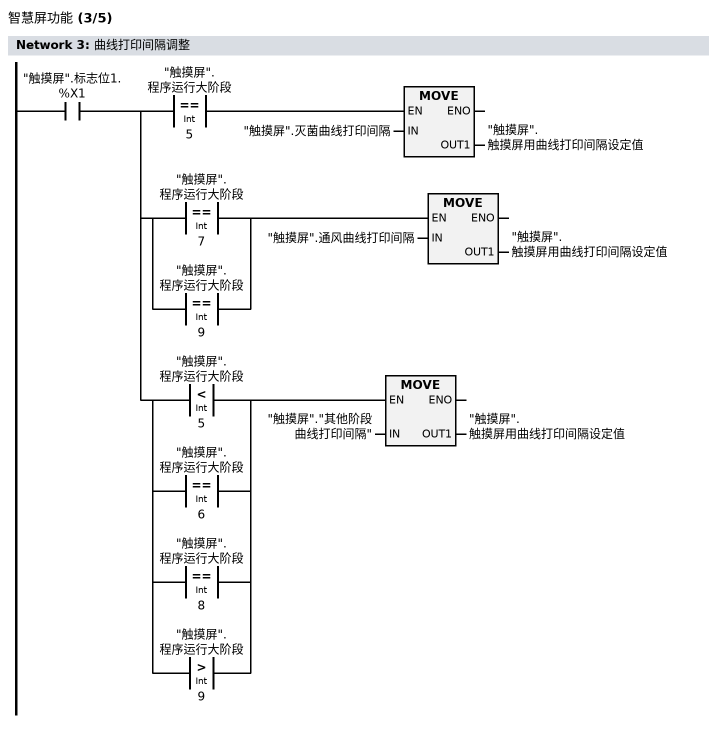
   RUNG wire#powerrail
      Contact( "触摸屏".标志位1.%X1 )
      wire#w1
      { S7_Templates := "SrcType := Int" } EQ_Contact(in1 := "触摸屏".程序运行大阶段, in2 := 5)
      Move(in := "触摸屏".灭菌曲线打印间隔, out1 => "触摸屏".触摸屏用曲线打印间隔设定值)
   END_RUNG
   RUNG wire#w1
      { S7_Templates := "SrcType := Int" } EQ_Contact(in1 := "触摸屏".程序运行大阶段, in2 := 7)
      wire#w2
      Move(in := "触摸屏".通风曲线打印间隔, out1 => "触摸屏".触摸屏用曲线打印间隔设定值)
   END_RUNG
   RUNG wire#w1
      { S7_Templates := "SrcType := Int" } EQ_Contact(in1 := "触摸屏".程序运行大阶段, in2 := 9)
   END_RUNG wire#w2
   RUNG wire#w1
      { S7_Templates := "SrcType := Int" } LT_Contact(in1 := "触摸屏".程序运行大阶段, in2 := 5)
      wire#w3
      Move(in := "触摸屏"."其他阶段 曲线打印间隔", out1 => "触摸屏".触摸屏用曲线打印间隔设定值)
   END_RUNG
   RUNG wire#w1
      { S7_Templates := "SrcType := Int" } EQ_Contact(in1 := "触摸屏".程序运行大阶段, in2 := 6)
   END_RUNG wire#w3
   RUNG wire#w1
      { S7_Templates := "SrcType := Int" } EQ_Contact(in1 := "触摸屏".程序运行大阶段, in2 := 8)
   END_RUNG wire#w3
   RUNG wire#w1
      { S7_Templates := "SrcType := Int" } GT_Contact(in1 := "触摸屏".程序运行大阶段, in2 := 9)
   END_RUNG wire#w3
   // the same network as SCL:
   IF "触摸屏".标志位1.%X1 AND ("触摸屏".程序运行大阶段 = 5) THEN "触摸屏".触摸屏用曲线打印间隔设定值 := "触摸屏".灭菌曲线打印间隔; END_IF;
   IF "触摸屏".标志位1.%X1 AND (("触摸屏".程序运行大阶段 = 7) OR ("触摸屏".程序运行大阶段 = 9)) THEN
       "触摸屏".触摸屏用曲线打印间隔设定值 := "触摸屏".通风曲线打印间隔;
   END_IF;
   IF "触摸屏".标志位1.%X1 AND (("触摸屏".程序运行大阶段 < 5) OR ("触摸屏".程序运行大阶段 = 6) OR ("触摸屏".程序运行大阶段 = 8) OR ("触摸屏".程序运行大阶段 > 9)) THEN
       "触摸屏".触摸屏用曲线打印间隔设定值 := "触摸屏"."其他阶段 曲线打印间隔";
   END_IF;
END_REGION

REGION Network 4: 报表打印控制 报表间隔控制，printflag， "DB48.DBD684", 用于控制报表打印
   // 曲线间隔：灭菌20秒，通风60秒，其他10秒
   // 报表间隔：1：预处理  10分钟
   // 2：保压   10分钟
   // 3：加湿    10分钟
   // 4：加药    10分钟
   // 5：灭菌    20分钟
   // 6：脉动    10分钟
   // 7：通风   60分钟
   // 8：紧急脉动 10分钟
   // 9：紧急通风  30分钟
   // 10：结束
   // 
   // 智慧屏曲线打印会打印：大阶段 小阶段  printflag+定时存储的数据，定时存储需要再global全局设置
   //             报表打印会打印：大阶段 小阶段  printflag
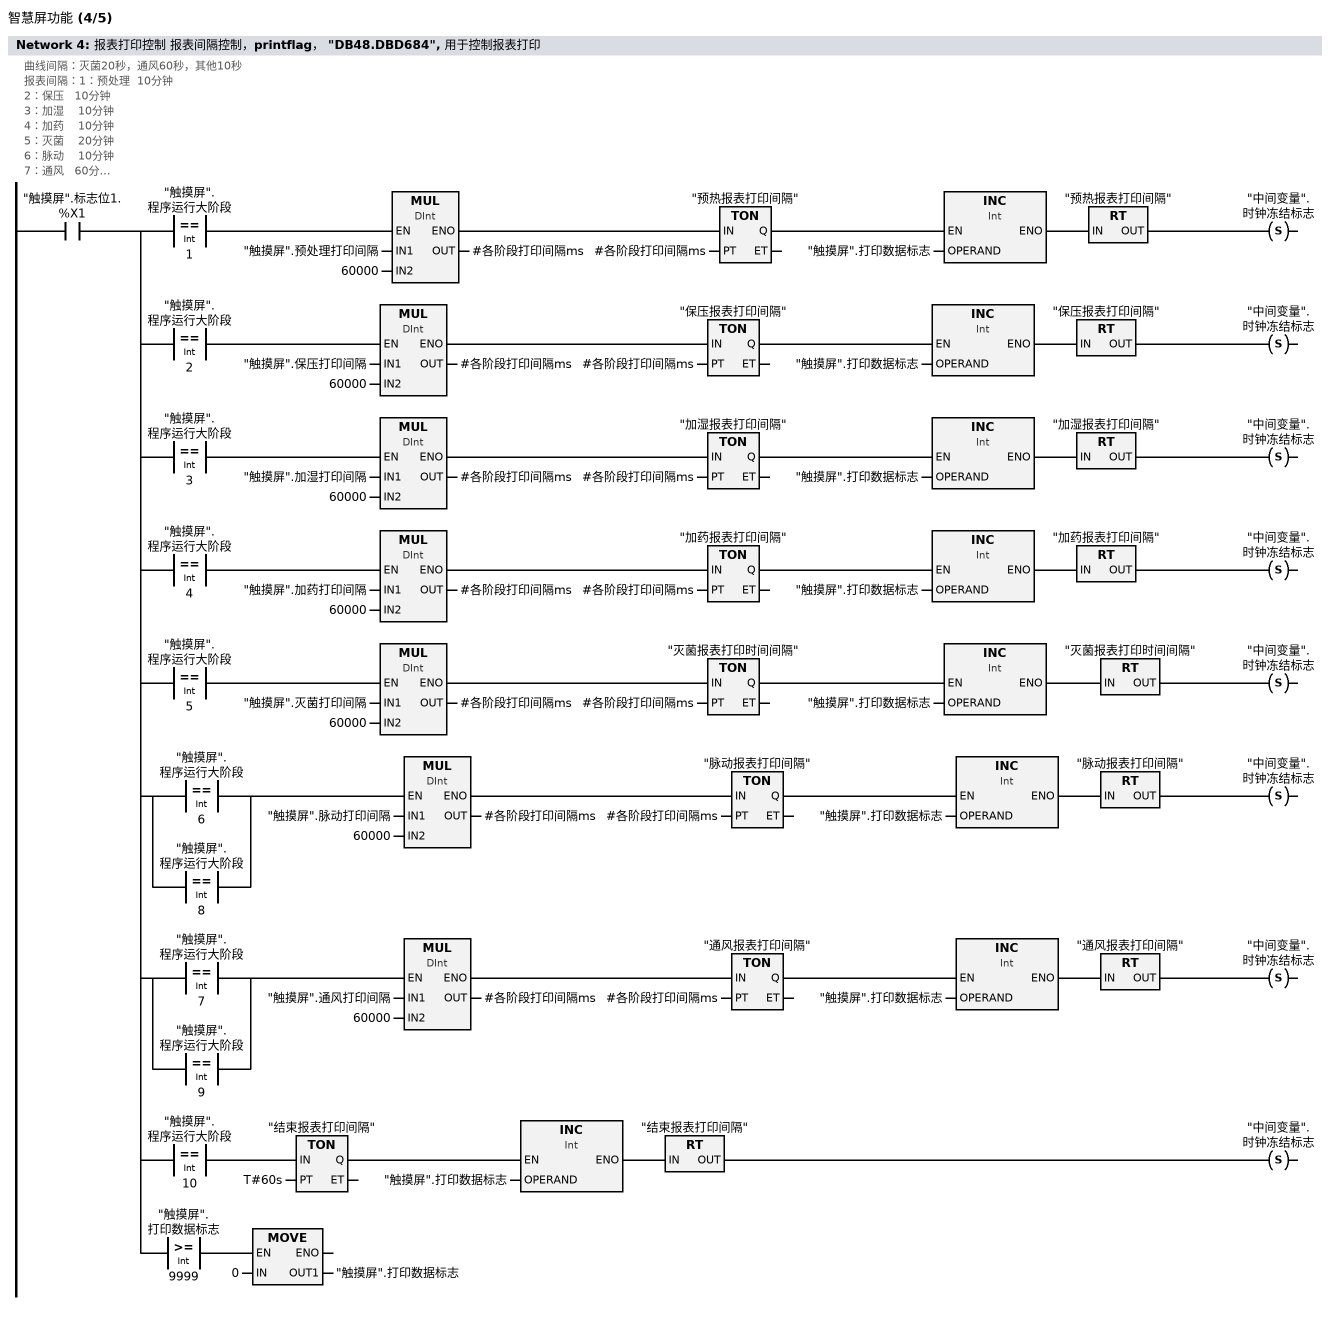
   #_w1 := "触摸屏".标志位1.%X1 AND ("触摸屏".程序运行大阶段 = 1);
   IF #_w1 THEN #各阶段打印间隔ms := "触摸屏".预处理打印间隔 * 60000; END_IF;
   "预热报表打印间隔".TON(IN := #_w1, PT := #各阶段打印间隔ms);
   IF "预热报表打印间隔".Q THEN "触摸屏".打印数据标志 := "触摸屏".打印数据标志 + 1; END_IF;
   #_w2 := "预热报表打印间隔".Q;
   IF #_w2 THEN
       RESET_TIMER("预热报表打印间隔");
       "中间变量".时钟冻结标志 := TRUE;
   END_IF;
   #_w3 := "触摸屏".标志位1.%X1 AND ("触摸屏".程序运行大阶段 = 2);
   IF #_w3 THEN #各阶段打印间隔ms := "触摸屏".保压打印间隔 * 60000; END_IF;
   "保压报表打印间隔".TON(IN := #_w3, PT := #各阶段打印间隔ms);
   IF "保压报表打印间隔".Q THEN "触摸屏".打印数据标志 := "触摸屏".打印数据标志 + 1; END_IF;
   #_w4 := "保压报表打印间隔".Q;
   IF #_w4 THEN
       RESET_TIMER("保压报表打印间隔");
       "中间变量".时钟冻结标志 := TRUE;
   END_IF;
   #_w5 := "触摸屏".标志位1.%X1 AND ("触摸屏".程序运行大阶段 = 3);
   IF #_w5 THEN #各阶段打印间隔ms := "触摸屏".加湿打印间隔 * 60000; END_IF;
   "加湿报表打印间隔".TON(IN := #_w5, PT := #各阶段打印间隔ms);
   IF "加湿报表打印间隔".Q THEN "触摸屏".打印数据标志 := "触摸屏".打印数据标志 + 1; END_IF;
   #_w6 := "加湿报表打印间隔".Q;
   IF #_w6 THEN
       RESET_TIMER("加湿报表打印间隔");
       "中间变量".时钟冻结标志 := TRUE;
   END_IF;
   #_w7 := "触摸屏".标志位1.%X1 AND ("触摸屏".程序运行大阶段 = 4);
   IF #_w7 THEN #各阶段打印间隔ms := "触摸屏".加药打印间隔 * 60000; END_IF;
   "加药报表打印间隔".TON(IN := #_w7, PT := #各阶段打印间隔ms);
   IF "加药报表打印间隔".Q THEN "触摸屏".打印数据标志 := "触摸屏".打印数据标志 + 1; END_IF;
   #_w8 := "加药报表打印间隔".Q;
   IF #_w8 THEN
       RESET_TIMER("加药报表打印间隔");
       "中间变量".时钟冻结标志 := TRUE;
   END_IF;
   #_w9 := "触摸屏".标志位1.%X1 AND ("触摸屏".程序运行大阶段 = 5);
   IF #_w9 THEN #各阶段打印间隔ms := "触摸屏".灭菌打印间隔 * 60000; END_IF;
   "灭菌报表打印时间间隔".TON(IN := #_w9, PT := #各阶段打印间隔ms);
   IF "灭菌报表打印时间间隔".Q THEN "触摸屏".打印数据标志 := "触摸屏".打印数据标志 + 1; END_IF;
   #_w10 := "灭菌报表打印时间间隔".Q;
   IF #_w10 THEN
       RESET_TIMER("灭菌报表打印时间间隔");
       "中间变量".时钟冻结标志 := TRUE;
   END_IF;
   #_w11 := "触摸屏".标志位1.%X1 AND (("触摸屏".程序运行大阶段 = 6) OR ("触摸屏".程序运行大阶段 = 8));
   IF #_w11 THEN #各阶段打印间隔ms := "触摸屏".脉动打印间隔 * 60000; END_IF;
   "脉动报表打印间隔".TON(IN := #_w11, PT := #各阶段打印间隔ms);
   IF "脉动报表打印间隔".Q THEN "触摸屏".打印数据标志 := "触摸屏".打印数据标志 + 1; END_IF;
   #_w12 := "脉动报表打印间隔".Q;
   IF #_w12 THEN
       RESET_TIMER("脉动报表打印间隔");
       "中间变量".时钟冻结标志 := TRUE;
   END_IF;
   #_w13 := "触摸屏".标志位1.%X1 AND (("触摸屏".程序运行大阶段 = 7) OR ("触摸屏".程序运行大阶段 = 9));
   IF #_w13 THEN #各阶段打印间隔ms := "触摸屏".通风打印间隔 * 60000; END_IF;
   "通风报表打印间隔".TON(IN := #_w13, PT := #各阶段打印间隔ms);
   IF "通风报表打印间隔".Q THEN "触摸屏".打印数据标志 := "触摸屏".打印数据标志 + 1; END_IF;
   #_w14 := "通风报表打印间隔".Q;
   IF #_w14 THEN
       RESET_TIMER("通风报表打印间隔");
       "中间变量".时钟冻结标志 := TRUE;
   END_IF;
   "结束报表打印间隔".TON(IN := "触摸屏".标志位1.%X1 AND ("触摸屏".程序运行大阶段 = 10), PT := T#60s);
   IF "结束报表打印间隔".Q THEN "触摸屏".打印数据标志 := "触摸屏".打印数据标志 + 1; END_IF;
   #_w15 := "结束报表打印间隔".Q;
   IF #_w15 THEN
       RESET_TIMER("结束报表打印间隔");
       "中间变量".时钟冻结标志 := TRUE;
   END_IF;
   IF "触摸屏".标志位1.%X1 AND ("触摸屏".打印数据标志 >= 9999) THEN "触摸屏".打印数据标志 := 0; END_IF;
END_REGION

REGION Network 5: 冻结PLC时钟标志，为了智慧屏能获取 阶段变化的真实时间，阶段变化后需要冻结PLC时间2秒钟
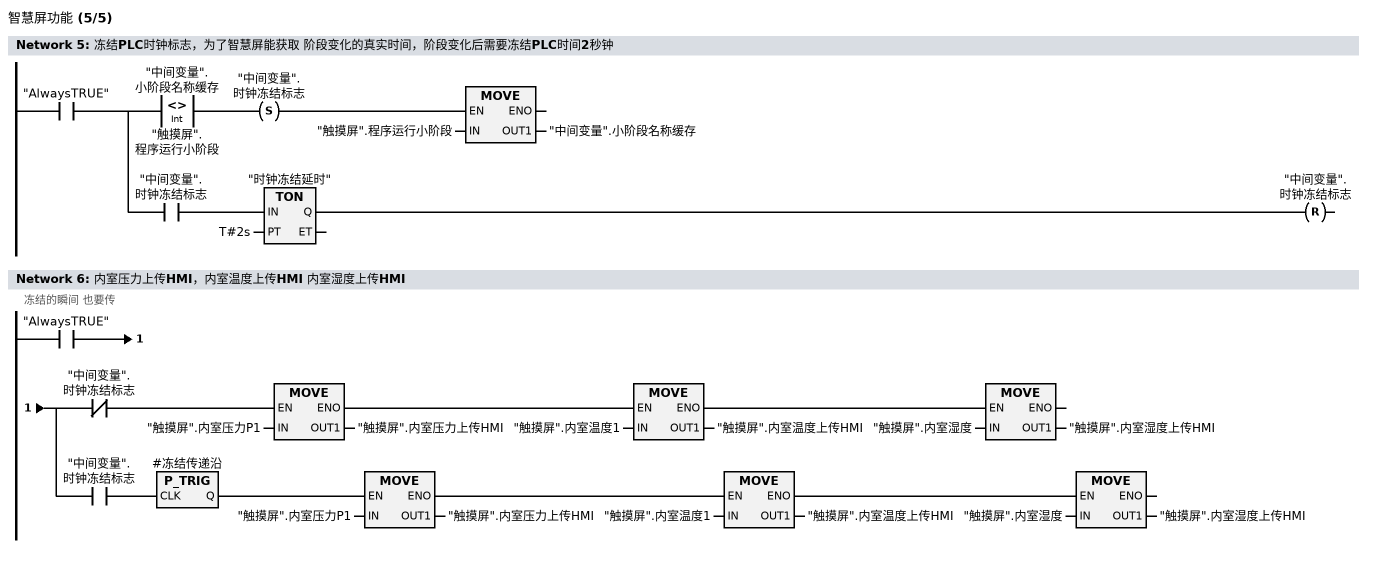
   IF "AlwaysTRUE" AND ("中间变量".小阶段名称缓存 <> "触摸屏".程序运行小阶段) THEN
       "中间变量".时钟冻结标志 := TRUE;
       "中间变量".小阶段名称缓存 := "触摸屏".程序运行小阶段;
   END_IF;
   "时钟冻结延时".TON(IN := "AlwaysTRUE" AND "中间变量".时钟冻结标志, PT := T#2s);
   IF "时钟冻结延时".Q THEN "中间变量".时钟冻结标志 := FALSE; END_IF;
END_REGION

REGION Network 6: 内室压力上传HMI，内室温度上传HMI 内室湿度上传HMI
   // 冻结的瞬间 也要传
   RUNG wire#powerrail
      Contact( "AlwaysTRUE" )
      wire#w1
      I_Contact( "中间变量".时钟冻结标志 )
      Move(in := "触摸屏".内室压力P1, out1 => "触摸屏".内室压力上传HMI)
      Move(in := "触摸屏".内室温度1, out1 => "触摸屏".内室温度上传HMI)
      Move(in := "触摸屏".内室湿度, out1 => "触摸屏".内室湿度上传HMI)
   END_RUNG
   RUNG wire#w1
      Contact( "中间变量".时钟冻结标志 )
      P_Trig( #冻结传递沿 )
      Move(in := "触摸屏".内室压力P1, out1 => "触摸屏".内室压力上传HMI)
      Move(in := "触摸屏".内室温度1, out1 => "触摸屏".内室温度上传HMI)
      Move(in := "触摸屏".内室湿度, out1 => "触摸屏".内室湿度上传HMI)
   END_RUNG
   // the same network as SCL:
   IF "AlwaysTRUE" AND NOT "中间变量".时钟冻结标志 THEN
       "触摸屏".内室压力上传HMI := "触摸屏".内室压力P1;
       "触摸屏".内室温度上传HMI := "触摸屏".内室温度1;
       "触摸屏".内室湿度上传HMI := "触摸屏".内室湿度;
   END_IF;
   #_w1 := "AlwaysTRUE" AND "中间变量".时钟冻结标志;
   #_w2 := #_w1 AND NOT #冻结传递沿;   // rising edge
   #冻结传递沿 := #_w1;
   IF #_w2 THEN
       "触摸屏".内室压力上传HMI := "触摸屏".内室压力P1;
       "触摸屏".内室温度上传HMI := "触摸屏".内室温度1;
       "触摸屏".内室湿度上传HMI := "触摸屏".内室湿度;
   END_IF;
END_REGION
END_FUNCTION_BLOCK

// folder: 6系统设置

FUNCTION_BLOCK "系统参数设置"   // FB21, LAD
{ S7_Optimized_Access := 'TRUE' }
VERSION : 0.1
   VAR
      催化剂使用时间秒 : Int;
      催化剂使用时间分 : Int;
      催化剂使用时间时 : Int;
      催化剂使用统计沿 : Bool;
   END_VAR
   VAR RETAIN
      催化剂使用统计秒 : Int;
   END_VAR
   VAR_TEMP
      中间变量 : Int;
   END_VAR
   VAR_TEMP   // added for the SCL form of the ladder/FBD networks
      _w1 : Bool;
      _w2 : Bool;
   END_VAR
BEGIN

REGION Network 1: 解毒阀开启时间统计，即催化剂使用时间统计
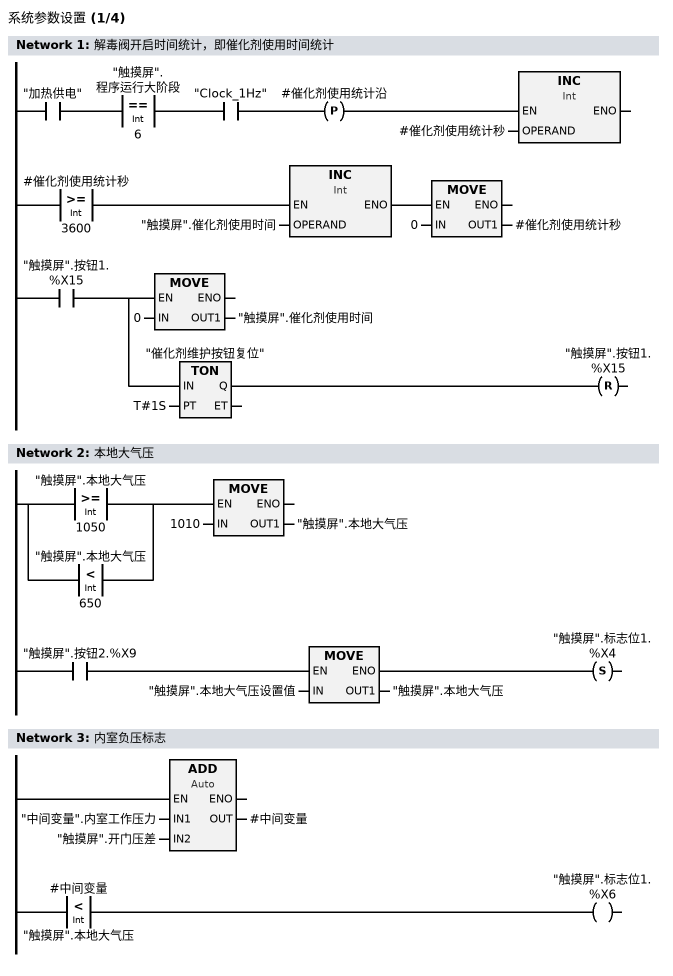
   #_w1 := "加热供电" AND ("触摸屏".程序运行大阶段 = 6) AND "Clock_1Hz";
   #_w2 := #_w1 AND NOT #催化剂使用统计沿;   // rising edge
   #催化剂使用统计沿 := #_w1;
   IF #_w2 THEN #催化剂使用统计秒 := #催化剂使用统计秒 + 1; END_IF;
   IF #催化剂使用统计秒 >= 3600 THEN
       "触摸屏".催化剂使用时间 := "触摸屏".催化剂使用时间 + 1;
       #催化剂使用统计秒 := 0;
   END_IF;
   IF "触摸屏".按钮1.%X15 THEN "触摸屏".催化剂使用时间 := 0; END_IF;
   "催化剂维护按钮复位".TON(IN := "触摸屏".按钮1.%X15, PT := T#1S);
   IF "催化剂维护按钮复位".Q THEN "触摸屏".按钮1.%X15 := FALSE; END_IF;
END_REGION

REGION Network 2: 本地大气压
   RUNG wire#powerrail
      { S7_Templates := "SrcType := Int" } GE_Contact(in1 := "触摸屏".本地大气压, in2 := 1050)
      wire#w1
      Move(in := 1010, out1 => "触摸屏".本地大气压)
   END_RUNG
   RUNG wire#powerrail
      { S7_Templates := "SrcType := Int" } LT_Contact(in1 := "触摸屏".本地大气压, in2 := 650)
   END_RUNG wire#w1
   RUNG wire#powerrail
      Contact( "触摸屏".按钮2.%X9 )
      Move(in := "触摸屏".本地大气压设置值, out1 => "触摸屏".本地大气压)
      S_Coil( "触摸屏".标志位1.%X4 )
   END_RUNG
   // the same network as SCL:
   IF ("触摸屏".本地大气压 >= 1050) OR ("触摸屏".本地大气压 < 650) THEN "触摸屏".本地大气压 := 1010; END_IF;
   IF "触摸屏".按钮2.%X9 THEN
       "触摸屏".本地大气压 := "触摸屏".本地大气压设置值;
       "触摸屏".标志位1.%X4 := TRUE;
   END_IF;
END_REGION

REGION Network 3: 内室负压标志
   RUNG wire#powerrail
      Add(in1 := "中间变量".内室工作压力, in2 := "触摸屏".开门压差, out => #中间变量)
   END_RUNG
   RUNG wire#powerrail
      { S7_Templates := "SrcType := Int" } LT_Contact(in1 := #中间变量, in2 := "触摸屏".本地大气压)
      Coil( "触摸屏".标志位1.%X6 )
   END_RUNG
   // the same network as SCL:
   #中间变量 := "中间变量".内室工作压力 + "触摸屏".开门压差;
   "触摸屏".标志位1.%X6 := #中间变量 < "触摸屏".本地大气压;
END_REGION

REGION Network 4: 蜂鸣器参数
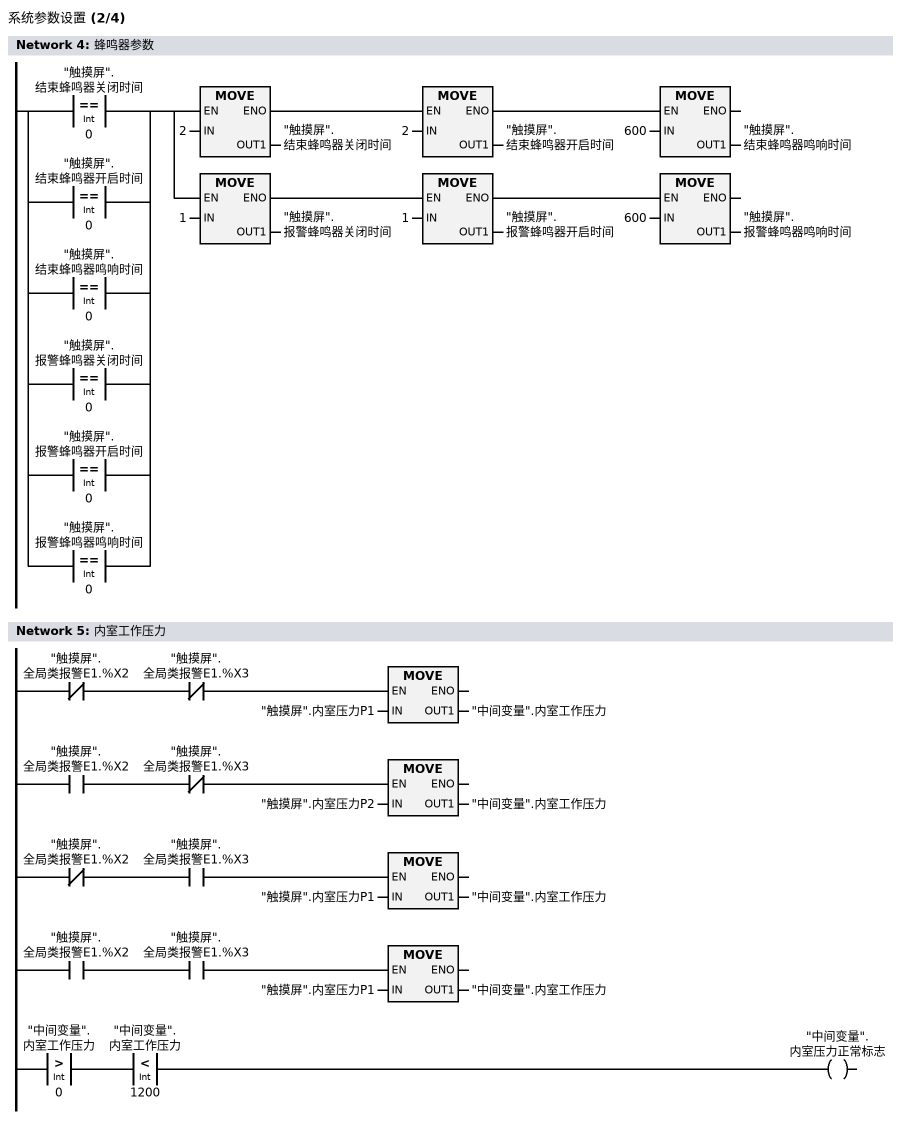
   RUNG wire#powerrail
      { S7_Templates := "SrcType := Int" } EQ_Contact(in1 := "触摸屏".结束蜂鸣器关闭时间, in2 := 0)
      wire#w1
      Move(in := 2, out1 => "触摸屏".结束蜂鸣器关闭时间)
      Move(in := 2, out1 => "触摸屏".结束蜂鸣器开启时间)
      Move(in := 600, out1 => "触摸屏".结束蜂鸣器鸣响时间)
   END_RUNG
   RUNG wire#powerrail
      { S7_Templates := "SrcType := Int" } EQ_Contact(in1 := "触摸屏".结束蜂鸣器开启时间, in2 := 0)
   END_RUNG wire#w1
   RUNG wire#powerrail
      { S7_Templates := "SrcType := Int" } EQ_Contact(in1 := "触摸屏".结束蜂鸣器鸣响时间, in2 := 0)
   END_RUNG wire#w1
   RUNG wire#powerrail
      { S7_Templates := "SrcType := Int" } EQ_Contact(in1 := "触摸屏".报警蜂鸣器关闭时间, in2 := 0)
   END_RUNG wire#w1
   RUNG wire#powerrail
      { S7_Templates := "SrcType := Int" } EQ_Contact(in1 := "触摸屏".报警蜂鸣器开启时间, in2 := 0)
   END_RUNG wire#w1
   RUNG wire#powerrail
      { S7_Templates := "SrcType := Int" } EQ_Contact(in1 := "触摸屏".报警蜂鸣器鸣响时间, in2 := 0)
   END_RUNG wire#w1
   RUNG wire#w1
      Move(in := 1, out1 => "触摸屏".报警蜂鸣器关闭时间)
      Move(in := 1, out1 => "触摸屏".报警蜂鸣器开启时间)
      Move(in := 600, out1 => "触摸屏".报警蜂鸣器鸣响时间)
   END_RUNG
   // the same network as SCL:
   #_w1 := ("触摸屏".结束蜂鸣器关闭时间 = 0) OR ("触摸屏".结束蜂鸣器开启时间 = 0) OR ("触摸屏".结束蜂鸣器鸣响时间 = 0) OR ("触摸屏".报警蜂鸣器关闭时间 = 0) OR ("触摸屏".报警蜂鸣器开启时间 = 0) OR ("触摸屏".报警蜂鸣器鸣响时间 = 0);
   #_w2 := ("触摸屏".结束蜂鸣器关闭时间 = 0) OR ("触摸屏".结束蜂鸣器开启时间 = 0) OR ("触摸屏".结束蜂鸣器鸣响时间 = 0) OR ("触摸屏".报警蜂鸣器关闭时间 = 0) OR ("触摸屏".报警蜂鸣器开启时间 = 0) OR ("触摸屏".报警蜂鸣器鸣响时间 = 0);
   IF #_w2 THEN
       "触摸屏".结束蜂鸣器关闭时间 := 2;
       "触摸屏".结束蜂鸣器开启时间 := 2;
       "触摸屏".结束蜂鸣器鸣响时间 := 600;
   END_IF;
   IF #_w1 THEN
       "触摸屏".报警蜂鸣器关闭时间 := 1;
       "触摸屏".报警蜂鸣器开启时间 := 1;
       "触摸屏".报警蜂鸣器鸣响时间 := 600;
   END_IF;
END_REGION

REGION Network 5: 内室工作压力
   RUNG wire#powerrail
      I_Contact( "触摸屏".全局类报警E1.%X2 )
      I_Contact( "触摸屏".全局类报警E1.%X3 )
      Move(in := "触摸屏".内室压力P1, out1 => "中间变量".内室工作压力)
   END_RUNG
   RUNG wire#powerrail
      Contact( "触摸屏".全局类报警E1.%X2 )
      I_Contact( "触摸屏".全局类报警E1.%X3 )
      Move(in := "触摸屏".内室压力P2, out1 => "中间变量".内室工作压力)
   END_RUNG
   RUNG wire#powerrail
      I_Contact( "触摸屏".全局类报警E1.%X2 )
      Contact( "触摸屏".全局类报警E1.%X3 )
      Move(in := "触摸屏".内室压力P1, out1 => "中间变量".内室工作压力)
   END_RUNG
   RUNG wire#powerrail
      Contact( "触摸屏".全局类报警E1.%X2 )
      Contact( "触摸屏".全局类报警E1.%X3 )
      Move(in := "触摸屏".内室压力P1, out1 => "中间变量".内室工作压力)
   END_RUNG
   RUNG wire#powerrail
      { S7_Templates := "SrcType := Int" } GT_Contact(in1 := "中间变量".内室工作压力, in2 := 0)
      { S7_Templates := "SrcType := Int" } LT_Contact(in1 := "中间变量".内室工作压力, in2 := 1200)
      Coil( "中间变量".内室压力正常标志 )
   END_RUNG
   // the same network as SCL:
   IF NOT "触摸屏".全局类报警E1.%X2 AND NOT "触摸屏".全局类报警E1.%X3 THEN "中间变量".内室工作压力 := "触摸屏".内室压力P1; END_IF;
   IF "触摸屏".全局类报警E1.%X2 AND NOT "触摸屏".全局类报警E1.%X3 THEN "中间变量".内室工作压力 := "触摸屏".内室压力P2; END_IF;
   IF NOT "触摸屏".全局类报警E1.%X2 AND "触摸屏".全局类报警E1.%X3 THEN "中间变量".内室工作压力 := "触摸屏".内室压力P1; END_IF;
   IF "触摸屏".全局类报警E1.%X2 AND "触摸屏".全局类报警E1.%X3 THEN "中间变量".内室工作压力 := "触摸屏".内室压力P1; END_IF;
   "中间变量".内室压力正常标志 := ("中间变量".内室工作压力 > 0) AND ("中间变量".内室工作压力 < 1200);
END_REGION

REGION Network 6: 设备维护
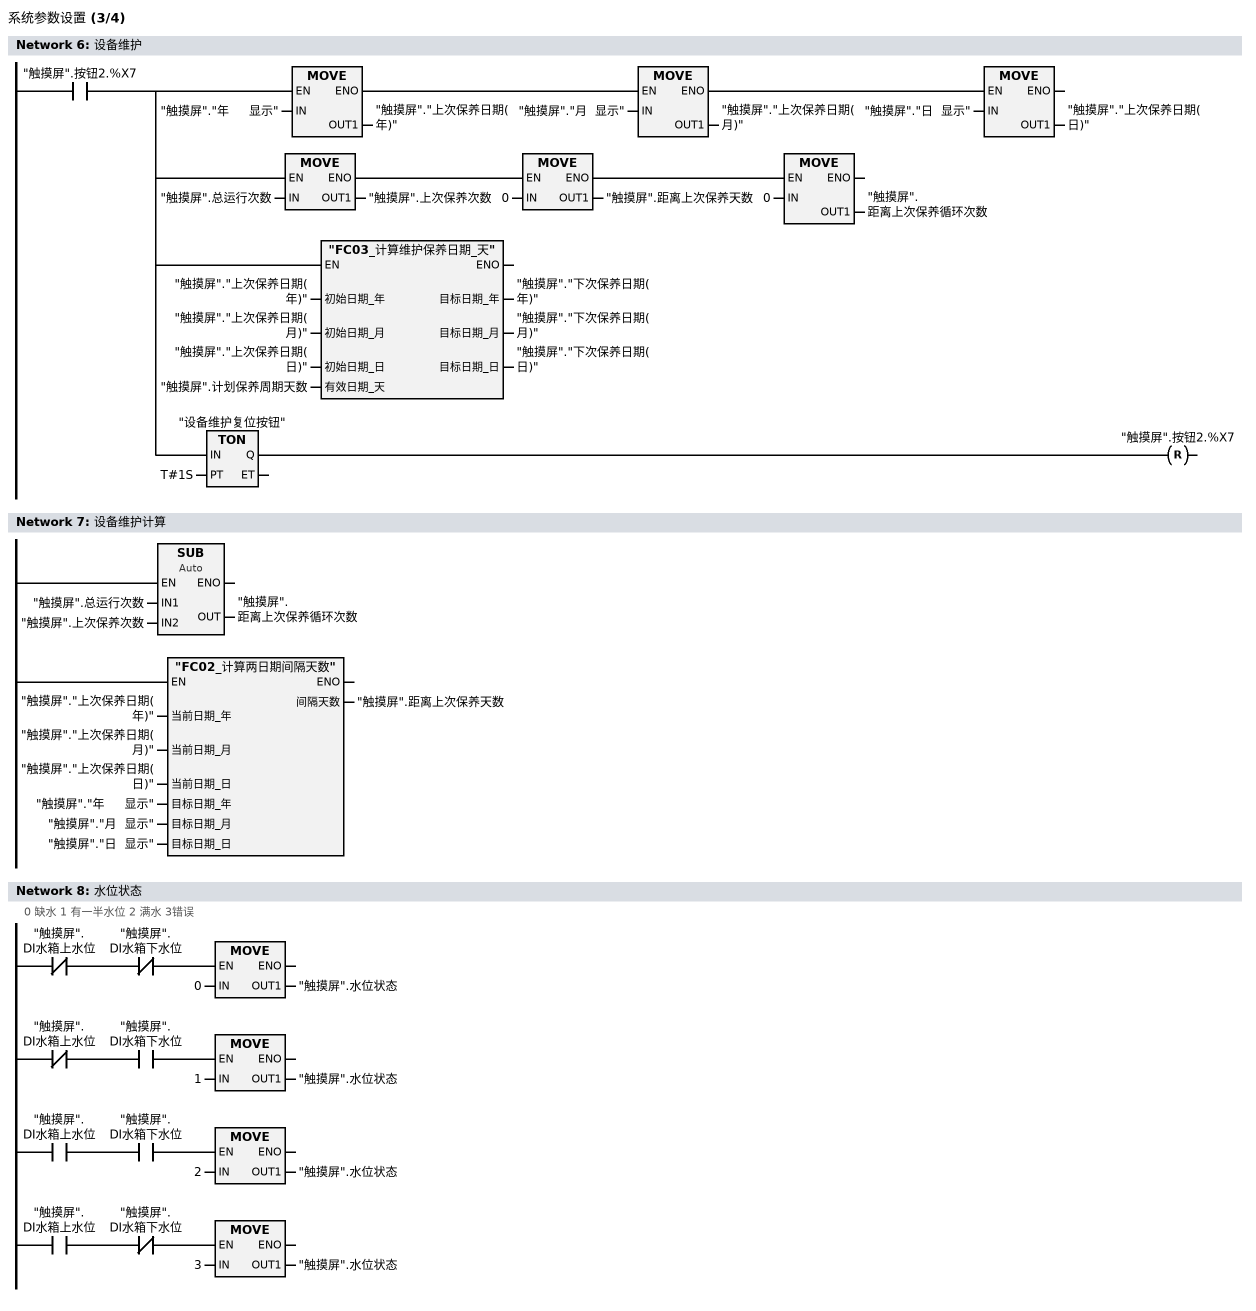
   IF "触摸屏".按钮2.%X7 THEN
       "触摸屏"."上次保养日期(年)" := "触摸屏"."年     显示";
       "触摸屏"."上次保养日期(月)" := "触摸屏"."月  显示";
       "触摸屏"."上次保养日期(日)" := "触摸屏"."日  显示";
       "触摸屏".上次保养次数 := "触摸屏".总运行次数;
       "触摸屏".距离上次保养天数 := 0;
       "触摸屏".距离上次保养循环次数 := 0;
   END_IF;
   #_w1 := "触摸屏".按钮2.%X7;
   IF #_w1 THEN
       "FC03_计算维护保养日期_天"(初始日期_年 := "触摸屏"."上次保养日期(年)",
                         初始日期_月 := "触摸屏"."上次保养日期(月)",
                         初始日期_日 := "触摸屏"."上次保养日期(日)",
                         有效日期_天 := "触摸屏".计划保养周期天数,
                         目标日期_年 => "触摸屏"."下次保养日期(年)",
                         目标日期_月 => "触摸屏"."下次保养日期(月)",
                         目标日期_日 => "触摸屏"."下次保养日期(日)");
   END_IF;
   "设备维护复位按钮".TON(IN := #_w1, PT := T#1S);
   IF "设备维护复位按钮".Q THEN "触摸屏".按钮2.%X7 := FALSE; END_IF;
END_REGION

REGION Network 7: 设备维护计算
   RUNG wire#powerrail
      Sub(in1 := "触摸屏".总运行次数, in2 := "触摸屏".上次保养次数, out => "触摸屏".距离上次保养循环次数)
   END_RUNG
   RUNG wire#powerrail
      "FC02_计算两日期间隔天数"(当前日期_年 := "触摸屏"."上次保养日期(年)", 当前日期_月 := "触摸屏"."上次保养日期(月)", 当前日期_日 := "触摸屏"."上次保养日期(日)", 目标日期_年 := "触摸屏"."年     显示", 目标日期_月 := "触摸屏"."月  显示", 目标日期_日 := "触摸屏"."日  显示", 间隔天数 => "触摸屏".距离上次保养天数)
   END_RUNG
   // the same network as SCL:
   "触摸屏".距离上次保养循环次数 := "触摸屏".总运行次数 - "触摸屏".上次保养次数;
   "FC02_计算两日期间隔天数"(当前日期_年 := "触摸屏"."上次保养日期(年)",
                    当前日期_月 := "触摸屏"."上次保养日期(月)",
                    当前日期_日 := "触摸屏"."上次保养日期(日)",
                    目标日期_年 := "触摸屏"."年     显示",
                    目标日期_月 := "触摸屏"."月  显示",
                    目标日期_日 := "触摸屏"."日  显示",
                    间隔天数 => "触摸屏".距离上次保养天数);
END_REGION

REGION Network 8: 水位状态
   // 0 缺水 1 有一半水位 2 满水 3错误
   RUNG wire#powerrail
      I_Contact( "触摸屏".DI水箱上水位 )
      I_Contact( "触摸屏".DI水箱下水位 )
      Move(in := 0, out1 => "触摸屏".水位状态)
   END_RUNG
   RUNG wire#powerrail
      I_Contact( "触摸屏".DI水箱上水位 )
      Contact( "触摸屏".DI水箱下水位 )
      Move(in := 1, out1 => "触摸屏".水位状态)
   END_RUNG
   RUNG wire#powerrail
      Contact( "触摸屏".DI水箱上水位 )
      Contact( "触摸屏".DI水箱下水位 )
      Move(in := 2, out1 => "触摸屏".水位状态)
   END_RUNG
   RUNG wire#powerrail
      Contact( "触摸屏".DI水箱上水位 )
      I_Contact( "触摸屏".DI水箱下水位 )
      Move(in := 3, out1 => "触摸屏".水位状态)
   END_RUNG
   // the same network as SCL:
   IF NOT "触摸屏".DI水箱上水位 AND NOT "触摸屏".DI水箱下水位 THEN "触摸屏".水位状态 := 0; END_IF;
   IF NOT "触摸屏".DI水箱上水位 AND "触摸屏".DI水箱下水位 THEN "触摸屏".水位状态 := 1; END_IF;
   IF "触摸屏".DI水箱上水位 AND "触摸屏".DI水箱下水位 THEN "触摸屏".水位状态 := 2; END_IF;
   IF "触摸屏".DI水箱上水位 AND NOT "触摸屏".DI水箱下水位 THEN "触摸屏".水位状态 := 3; END_IF;
END_REGION

REGION Network 9: 气罐状态（66256中的是否扫描，是否更换没处理）
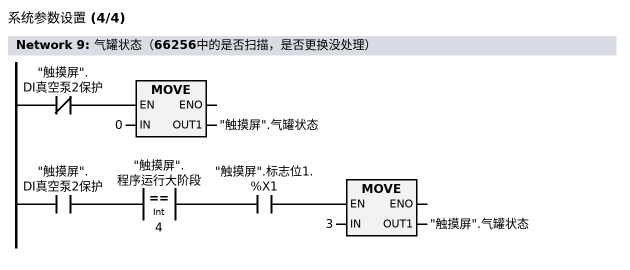
   RUNG wire#powerrail
      I_Contact( "触摸屏".DI真空泵2保护 )
      Move(in := 0, out1 => "触摸屏".气罐状态)
   END_RUNG
   RUNG wire#powerrail
      Contact( "触摸屏".DI真空泵2保护 )
      { S7_Templates := "SrcType := Int" } EQ_Contact(in1 := "触摸屏".程序运行大阶段, in2 := 4)
      Contact( "触摸屏".标志位1.%X1 )
      Move(in := 3, out1 => "触摸屏".气罐状态)
   END_RUNG
   // the same network as SCL:
   IF NOT "触摸屏".DI真空泵2保护 THEN "触摸屏".气罐状态 := 0; END_IF;
   IF "触摸屏".DI真空泵2保护 AND ("触摸屏".程序运行大阶段 = 4) AND "触摸屏".标志位1.%X1 THEN "触摸屏".气罐状态 := 3; END_IF;
END_REGION
END_FUNCTION_BLOCK

FUNCTION "FC02_计算两日期间隔天数" : Void   // FC9, SCL
{ S7_Optimized_Access := 'TRUE' }
VERSION : 0.1
   VAR_INPUT
      当前日期_年 : Int;
      当前日期_月 : Int;
      当前日期_日 : Int;
      目标日期_年 : Int;
      目标日期_月 : Int;
      目标日期_日 : Int;
   END_VAR
   VAR_OUTPUT
      间隔天数 : Int;
   END_VAR
   VAR_TEMP
      temp1 : Array[0..2] of Int;
      temp2 : Array[0..2] of Int;
   END_VAR
BEGIN
   (*
   算法解析：
   该算法总体思想是计算给定日期到公元元年3月1日的天数，然后相减，获取天数的间隔。
   m1 = (month_start + 9) % 12
   用于判断日期是否大于3月（2月是判断闰年的标识），还用于纪录到3月的间隔月数。
   y1 = year_start - m1/10
   判断如果是1月和2月，则不包括当前年（因为是计算到0年3月1日的天数）。
   d1 = 365*y1 + y1/4 - y1/100 + y1/400 + (m1*306 + 5)/10 + (day_start - 1)
   其中 365*y1 是不算闰年多出那一天的天数。
   y1/4 - y1/100 + y1/400
   是加所有闰年多出的那一天，四年一润，百年不润，四百年再润。
   (m2*306 + 5)/10
   用于计算到当前月到3月1日间的天数，306=365-31-28（1月和2月）
   5是全年中不是31天月份的个数，【31、28/29、31、30、31、30、31、31、30、31、30、31】。
   (day_start - 1)
   用于计算当前日到1日的间隔天数。
   *)
   #temp1[0] := (#当前日期_月 + 9) MOD 12;
   #temp1[1] := #当前日期_年 - #temp1[0] / 10;
   #temp1[2] := #temp1[1] * 365 + #temp1[1] / 4 - #temp1[1] / 100 + #temp1[1] / 400 + (#temp1[0] * 306 + 5) / 10 + (#当前日期_日 - 1);
   //IN1* 365+ IN1/4-IN1/ 100+IN1/400+ (IN2*306+5)/10+ (IN3-1)
   #temp2[0] := (#目标日期_月 + 9) MOD 12;
   #temp2[1] := #目标日期_年 - #temp2[0] / 10;
   #temp2[2] := #temp2[1] * 365 + #temp2[1] / 4 - #temp2[1] / 100 + #temp2[1] / 400 + (#temp2[0] * 306 + 5) / 10 + (#目标日期_日 - 1);
   #间隔天数 := #temp2[2] - #temp1[2];
   IF #间隔天数 < 0 THEN
       #间隔天数 := 0;

   END_IF;
END_FUNCTION

FUNCTION "FC03_计算维护保养日期_天" : Void   // FC10, SCL
{ S7_Optimized_Access := 'TRUE' }
VERSION : 0.1
   VAR_INPUT
      初始日期_年 : UInt;
      初始日期_月 : USInt;
      初始日期_日 : USInt;
      有效日期_天 : DInt;
   END_VAR
   VAR_OUTPUT
      目标日期_年 : UInt;
      目标日期_月 : USInt;
      目标日期_日 : USInt;
   END_VAR
   VAR_TEMP
      I : Int;
      N_年 : UInt;
      N_月 : USInt;
      N_日 : USInt;
      目标天数 : DInt;
      N月 : Array[0..12] of USInt;
   END_VAR
BEGIN
   //写入初始日期
   #N_年 := #初始日期_年;
   #N_月 := #初始日期_月;
   #N_日 := #初始日期_日;
   #目标天数 := #有效日期_天;
   //初始化每个月的日期
   FOR #I := 1 TO 12 DO
       CASE #I OF
           1, 3, 5, 7, 8, 10, 12:
               #N月[#I] := 31;
           4, 6, 9, 11:
               #N月[#I] := 30;
           ELSE
               #N月[#I] := 28;
       END_CASE;
   END_FOR;
   //闰年2月天数判断
   IF (#N_年 MOD 4 = 0) AND (#N_年 / 400 <> 0) OR (#N_年 / 400 = 0) THEN
       #N月[2] := 29;
   ELSE
       #N月[2] := 28;
   END_IF;
   //判断否跨月
   WHILE #目标天数 > (#N月[#N_月] - #N_日) DO
       #目标天数 := #目标天数 - (#N月[#N_月] - #N_日);
       #N_日 := 0;
       #N_月 := #N_月 + 1;
       //跨月后判断是否跨年
       IF #N_月 = 13 THEN
           #N_年 := #N_年 + 1;
           #N_月 := 1;
           IF (#N_年 MOD 4 = 0) AND (#N_年 / 400 <> 0) OR (#N_年 / 400 = 0) THEN
               #N月[2] := 29;
           ELSE
               #N月[2] := 28;
           END_IF;
       END_IF;
   END_WHILE;
   #目标日期_年 := #N_年;
   #目标日期_月 := #N_月;
   #目标日期_日 := DINT_TO_USINT(#目标天数 + #N_日);
END_FUNCTION

// folder: 7程序参数

FUNCTION_BLOCK "参数恢复默认"   // FB1, LAD
{ S7_Optimized_Access := 'TRUE' }
VERSION : 0.1
   VAR
      沿1 : Bool;
      沿2 : Bool;
      沿3 : Bool;
      沿4 : Bool;
      沿5 : Bool;
      沿6 : Bool;
      沿7 : Bool;
   END_VAR
   VAR_TEMP   // added for the SCL form of the ladder/FBD networks
      _w1 : Bool;
      _w2 : Bool;
      _w3 : Bool;
   END_VAR
BEGIN

REGION Network 1: 37℃程序参数恢复默认
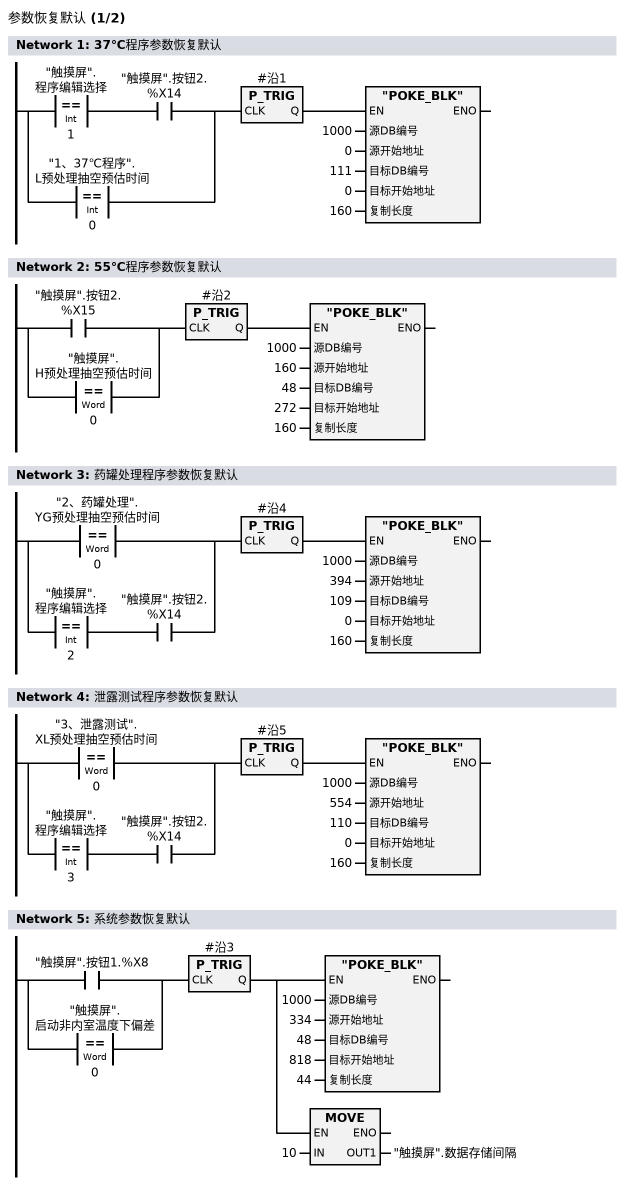
   RUNG wire#powerrail
      { S7_Templates := "SrcType := Int" } EQ_Contact(in1 := "触摸屏".程序编辑选择, in2 := 1)
      Contact( "触摸屏".按钮2.%X14 )
      wire#w1
      P_Trig( #沿1 )
      "POKE_BLK"(源DB编号 := 1000, 源开始地址 := 0, 目标DB编号 := 111, 目标开始地址 := 0, 复制长度 := 160)
   END_RUNG
   RUNG wire#powerrail
      { S7_Templates := "SrcType := Int" } EQ_Contact(in1 := "1、37℃程序".L预处理抽空预估时间, in2 := 0)
   END_RUNG wire#w1
   // the same network as SCL:
   #_w1 := (("触摸屏".程序编辑选择 = 1) AND "触摸屏".按钮2.%X14) OR ("1、37℃程序".L预处理抽空预估时间 = 0);
   #_w2 := #_w1 AND NOT #沿1;   // rising edge
   #沿1 := #_w1;
   IF #_w2 THEN "POKE_BLK"(源DB编号 := 1000, 源开始地址 := 0, 目标DB编号 := 111, 目标开始地址 := 0, 复制长度 := 160); END_IF;
END_REGION

REGION Network 2: 55℃程序参数恢复默认
   RUNG wire#powerrail
      Contact( "触摸屏".按钮2.%X15 )
      wire#w1
      P_Trig( #沿2 )
      "POKE_BLK"(源DB编号 := 1000, 源开始地址 := 160, 目标DB编号 := 48, 目标开始地址 := 272, 复制长度 := 160)
   END_RUNG
   RUNG wire#powerrail
      { S7_Templates := "SrcType := Word" } EQ_Contact(in1 := "触摸屏".H预处理抽空预估时间, in2 := 0)
   END_RUNG wire#w1
   // the same network as SCL:
   #_w1 := "触摸屏".按钮2.%X15 OR ("触摸屏".H预处理抽空预估时间 = 0);
   #_w2 := #_w1 AND NOT #沿2;   // rising edge
   #沿2 := #_w1;
   IF #_w2 THEN "POKE_BLK"(源DB编号 := 1000, 源开始地址 := 160, 目标DB编号 := 48, 目标开始地址 := 272, 复制长度 := 160); END_IF;
END_REGION

REGION Network 3: 药罐处理程序参数恢复默认
   RUNG wire#powerrail
      { S7_Templates := "SrcType := Word" } EQ_Contact(in1 := "2、药罐处理".YG预处理抽空预估时间, in2 := 0)
      wire#w1
      P_Trig( #沿4 )
      "POKE_BLK"(源DB编号 := 1000, 源开始地址 := 394, 目标DB编号 := 109, 目标开始地址 := 0, 复制长度 := 160)
   END_RUNG
   RUNG wire#powerrail
      { S7_Templates := "SrcType := Int" } EQ_Contact(in1 := "触摸屏".程序编辑选择, in2 := 2)
      Contact( "触摸屏".按钮2.%X14 )
   END_RUNG wire#w1
   // the same network as SCL:
   #_w1 := ("2、药罐处理".YG预处理抽空预估时间 = 0) OR (("触摸屏".程序编辑选择 = 2) AND "触摸屏".按钮2.%X14);
   #_w2 := #_w1 AND NOT #沿4;   // rising edge
   #沿4 := #_w1;
   IF #_w2 THEN "POKE_BLK"(源DB编号 := 1000, 源开始地址 := 394, 目标DB编号 := 109, 目标开始地址 := 0, 复制长度 := 160); END_IF;
END_REGION

REGION Network 4: 泄露测试程序参数恢复默认
   RUNG wire#powerrail
      { S7_Templates := "SrcType := Word" } EQ_Contact(in1 := "3、泄露测试".XL预处理抽空预估时间, in2 := 0)
      wire#w1
      P_Trig( #沿5 )
      "POKE_BLK"(源DB编号 := 1000, 源开始地址 := 554, 目标DB编号 := 110, 目标开始地址 := 0, 复制长度 := 160)
   END_RUNG
   RUNG wire#powerrail
      { S7_Templates := "SrcType := Int" } EQ_Contact(in1 := "触摸屏".程序编辑选择, in2 := 3)
      Contact( "触摸屏".按钮2.%X14 )
   END_RUNG wire#w1
   // the same network as SCL:
   #_w1 := ("3、泄露测试".XL预处理抽空预估时间 = 0) OR (("触摸屏".程序编辑选择 = 3) AND "触摸屏".按钮2.%X14);
   #_w2 := #_w1 AND NOT #沿5;   // rising edge
   #沿5 := #_w1;
   IF #_w2 THEN "POKE_BLK"(源DB编号 := 1000, 源开始地址 := 554, 目标DB编号 := 110, 目标开始地址 := 0, 复制长度 := 160); END_IF;
END_REGION

REGION Network 5: 系统参数恢复默认
   RUNG wire#powerrail
      Contact( "触摸屏".按钮1.%X8 )
      wire#w1
      P_Trig( #沿3 )
      wire#w2
      "POKE_BLK"(源DB编号 := 1000, 源开始地址 := 334, 目标DB编号 := 48, 目标开始地址 := 818, 复制长度 := 44)
   END_RUNG
   RUNG wire#powerrail
      { S7_Templates := "SrcType := Word" } EQ_Contact(in1 := "触摸屏".启动非内室温度下偏差, in2 := 0)
   END_RUNG wire#w1
   RUNG wire#w2
      { S7_GenerateENO := "TRUE" } Move(in := 10, out1 => "触摸屏".数据存储间隔)
   END_RUNG
   // the same network as SCL:
   #_w1 := "触摸屏".按钮1.%X8 OR ("触摸屏".启动非内室温度下偏差 = 0);
   #_w2 := #_w1 AND NOT #沿3;   // rising edge
   #沿3 := #_w1;
   IF #_w2 THEN
       "POKE_BLK"(源DB编号 := 1000, 源开始地址 := 334, 目标DB编号 := 48, 目标开始地址 := 818, 复制长度 := 44);
       "触摸屏".数据存储间隔 := 10;
   END_IF;
END_REGION

REGION Network 6: 偏差校准恢复默认
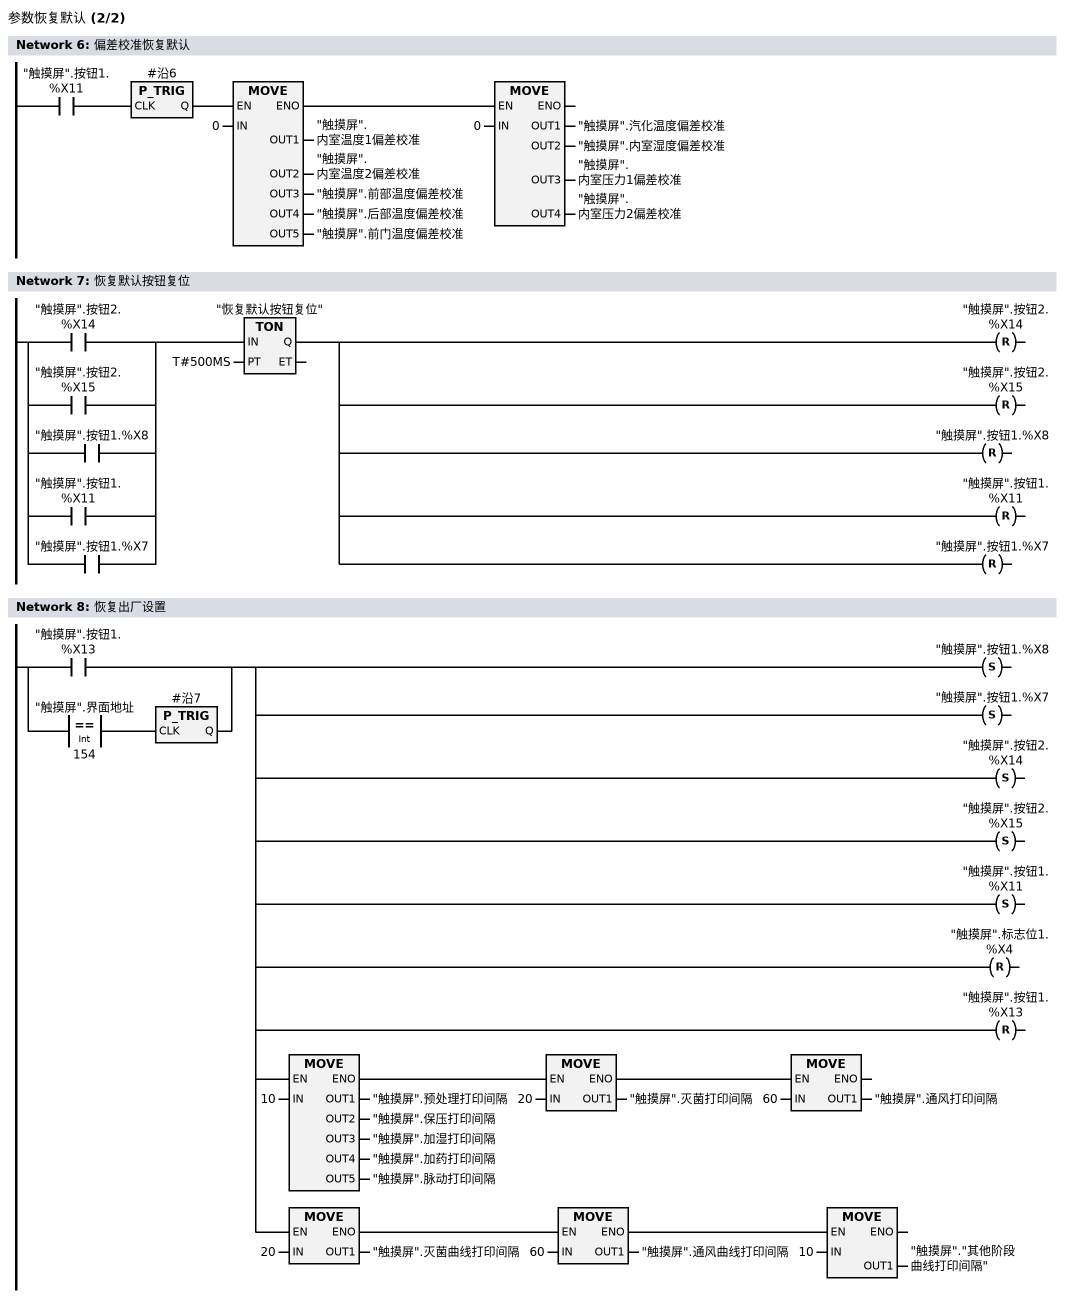
   RUNG wire#powerrail
      Contact( "触摸屏".按钮1.%X11 )
      P_Trig( #沿6 )
      Move(in := 0, out1 => "触摸屏".内室温度1偏差校准, out2 => "触摸屏".内室温度2偏差校准, out3 => "触摸屏".前部温度偏差校准, out4 => "触摸屏".后部温度偏差校准, out5 => "触摸屏".前门温度偏差校准)
      Move(in := 0, out1 => "触摸屏".汽化温度偏差校准, out2 => "触摸屏".内室湿度偏差校准, out3 => "触摸屏".内室压力1偏差校准, out4 => "触摸屏".内室压力2偏差校准)
   END_RUNG
   // the same network as SCL:
   #_w1 := "触摸屏".按钮1.%X11 AND NOT #沿6;   // rising edge
   #沿6 := "触摸屏".按钮1.%X11;
   IF #_w1 THEN
       "触摸屏".内室温度1偏差校准 := 0;
       "触摸屏".内室温度2偏差校准 := 0;
       "触摸屏".前部温度偏差校准 := 0;
       "触摸屏".后部温度偏差校准 := 0;
       "触摸屏".前门温度偏差校准 := 0;
       "触摸屏".汽化温度偏差校准 := 0;
       "触摸屏".内室湿度偏差校准 := 0;
       "触摸屏".内室压力1偏差校准 := 0;
       "触摸屏".内室压力2偏差校准 := 0;
   END_IF;
END_REGION

REGION Network 7: 恢复默认按钮复位
   "恢复默认按钮复位".TON(IN := "触摸屏".按钮2.%X14 OR "触摸屏".按钮2.%X15 OR "触摸屏".按钮1.%X8 OR "触摸屏".按钮1.%X11 OR "触摸屏".按钮1.%X7,
                  PT := T#500MS);
   IF "恢复默认按钮复位".Q THEN
       "触摸屏".按钮2.%X14 := FALSE;
       "触摸屏".按钮2.%X15 := FALSE;
       "触摸屏".按钮1.%X8 := FALSE;
       "触摸屏".按钮1.%X11 := FALSE;
       "触摸屏".按钮1.%X7 := FALSE;
   END_IF;
END_REGION

REGION Network 8: 恢复出厂设置
   RUNG wire#powerrail
      Contact( "触摸屏".按钮1.%X13 )
      wire#w1
      S_Coil( "触摸屏".按钮1.%X8 )
   END_RUNG
   RUNG wire#powerrail
      { S7_Templates := "SrcType := Int" } EQ_Contact(in1 := "触摸屏".界面地址, in2 := 154)
      P_Trig( #沿7 )
   END_RUNG wire#w1
   RUNG wire#w1
      S_Coil( "触摸屏".按钮1.%X7 )
   END_RUNG
   RUNG wire#w1
      S_Coil( "触摸屏".按钮2.%X14 )
   END_RUNG
   RUNG wire#w1
      S_Coil( "触摸屏".按钮2.%X15 )
   END_RUNG
   RUNG wire#w1
      S_Coil( "触摸屏".按钮1.%X11 )
   END_RUNG
   RUNG wire#w1
      R_Coil( "触摸屏".标志位1.%X4 )
   END_RUNG
   RUNG wire#w1
      R_Coil( "触摸屏".按钮1.%X13 )
   END_RUNG
   RUNG wire#w1
      Move(in := 10, out1 => "触摸屏".预处理打印间隔, out2 => "触摸屏".保压打印间隔, out3 => "触摸屏".加湿打印间隔, out4 => "触摸屏".加药打印间隔, out5 => "触摸屏".脉动打印间隔)
      Move(in := 20, out1 => "触摸屏".灭菌打印间隔)
      Move(in := 60, out1 => "触摸屏".通风打印间隔)
   END_RUNG
   RUNG wire#w1
      Move(in := 20, out1 => "触摸屏".灭菌曲线打印间隔)
      Move(in := 60, out1 => "触摸屏".通风曲线打印间隔)
      Move(in := 10, out1 => "触摸屏"."其他阶段 曲线打印间隔")
   END_RUNG
   // the same network as SCL:
   #_w1 := "触摸屏".界面地址 = 154;
   #_w2 := #_w1 AND NOT #沿7;   // rising edge
   #沿7 := #_w1;
   #_w3 := "触摸屏".按钮1.%X13 OR #_w2;
   IF #_w3 THEN
       "触摸屏".按钮1.%X8 := TRUE;
       "触摸屏".按钮1.%X7 := TRUE;
       "触摸屏".按钮2.%X14 := TRUE;
       "触摸屏".按钮2.%X15 := TRUE;
       "触摸屏".按钮1.%X11 := TRUE;
       "触摸屏".标志位1.%X4 := FALSE;
       "触摸屏".按钮1.%X13 := FALSE;
       "触摸屏".预处理打印间隔 := 10;
       "触摸屏".保压打印间隔 := 10;
       "触摸屏".加湿打印间隔 := 10;
       "触摸屏".加药打印间隔 := 10;
       "触摸屏".脉动打印间隔 := 10;
       "触摸屏".灭菌打印间隔 := 20;
       "触摸屏".通风打印间隔 := 60;
       "触摸屏".灭菌曲线打印间隔 := 20;
       "触摸屏".通风曲线打印间隔 := 60;
       "触摸屏"."其他阶段 曲线打印间隔" := 10;
   END_IF;
END_REGION
END_FUNCTION_BLOCK

FUNCTION_BLOCK "程序运行参数传递"   // FB2, LAD
{ S7_Optimized_Access := 'TRUE' }
VERSION : 0.1
   VAR
      沿1 : Bool;
      沿2 : Bool;
      沿3 : Bool;
      沿4 : Bool;
      沿5 : Bool;
      沿6 : Bool;
      沿7 : Bool;
   END_VAR
   VAR_TEMP   // added for the SCL form of the ladder/FBD networks
      _w1 : Bool;
   END_VAR
BEGIN

REGION Network 1: 37℃程序参数传递
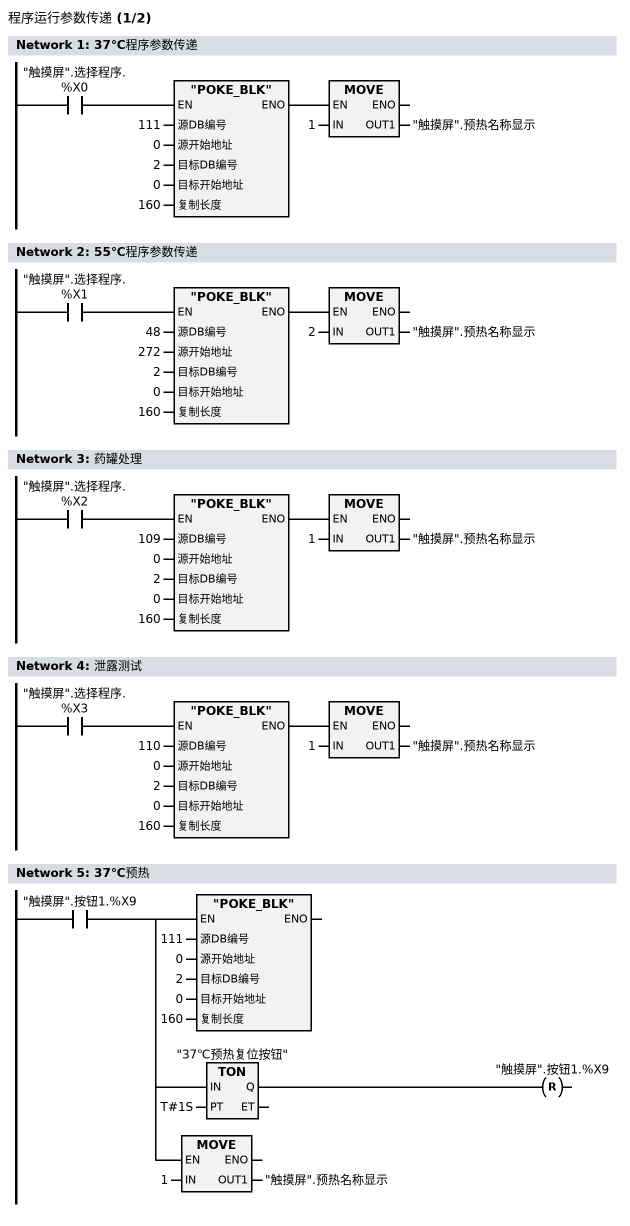
   RUNG wire#powerrail
      Contact( "触摸屏".选择程序.%X0 )
      "POKE_BLK"(源DB编号 := 111, 源开始地址 := 0, 目标DB编号 := 2, 目标开始地址 := 0, 复制长度 := 160)
      Move(in := 1, out1 => "触摸屏".预热名称显示)
   END_RUNG
   // the same network as SCL:
   "POKE_BLK"(EN := "触摸屏".选择程序.%X0,
              源DB编号 := 111,
              源开始地址 := 0,
              目标DB编号 := 2,
              目标开始地址 := 0,
              复制长度 := 160,
              ENO => #_w1);
   IF #_w1 THEN "触摸屏".预热名称显示 := 1; END_IF;
END_REGION

REGION Network 2: 55℃程序参数传递
   RUNG wire#powerrail
      Contact( "触摸屏".选择程序.%X1 )
      "POKE_BLK"(源DB编号 := 48, 源开始地址 := 272, 目标DB编号 := 2, 目标开始地址 := 0, 复制长度 := 160)
      Move(in := 2, out1 => "触摸屏".预热名称显示)
   END_RUNG
   // the same network as SCL:
   "POKE_BLK"(EN := "触摸屏".选择程序.%X1,
              源DB编号 := 48,
              源开始地址 := 272,
              目标DB编号 := 2,
              目标开始地址 := 0,
              复制长度 := 160,
              ENO => #_w1);
   IF #_w1 THEN "触摸屏".预热名称显示 := 2; END_IF;
END_REGION

REGION Network 3: 药罐处理
   RUNG wire#powerrail
      Contact( "触摸屏".选择程序.%X2 )
      "POKE_BLK"(源DB编号 := 109, 源开始地址 := 0, 目标DB编号 := 2, 目标开始地址 := 0, 复制长度 := 160)
      Move(in := 1, out1 => "触摸屏".预热名称显示)
   END_RUNG
   // the same network as SCL:
   "POKE_BLK"(EN := "触摸屏".选择程序.%X2,
              源DB编号 := 109,
              源开始地址 := 0,
              目标DB编号 := 2,
              目标开始地址 := 0,
              复制长度 := 160,
              ENO => #_w1);
   IF #_w1 THEN "触摸屏".预热名称显示 := 1; END_IF;
END_REGION

REGION Network 4: 泄露测试
   RUNG wire#powerrail
      Contact( "触摸屏".选择程序.%X3 )
      "POKE_BLK"(源DB编号 := 110, 源开始地址 := 0, 目标DB编号 := 2, 目标开始地址 := 0, 复制长度 := 160)
      Move(in := 1, out1 => "触摸屏".预热名称显示)
   END_RUNG
   // the same network as SCL:
   "POKE_BLK"(EN := "触摸屏".选择程序.%X3,
              源DB编号 := 110,
              源开始地址 := 0,
              目标DB编号 := 2,
              目标开始地址 := 0,
              复制长度 := 160,
              ENO => #_w1);
   IF #_w1 THEN "触摸屏".预热名称显示 := 1; END_IF;
END_REGION

REGION Network 5: 37℃预热
   #_w1 := "触摸屏".按钮1.%X9;
   IF #_w1 THEN "POKE_BLK"(源DB编号 := 111, 源开始地址 := 0, 目标DB编号 := 2, 目标开始地址 := 0, 复制长度 := 160); END_IF;
   "37℃预热复位按钮".TON(IN := #_w1, PT := T#1S);
   IF "37℃预热复位按钮".Q THEN "触摸屏".按钮1.%X9 := FALSE; END_IF;
   IF #_w1 THEN "触摸屏".预热名称显示 := 1; END_IF;
END_REGION

REGION Network 6: 55℃预热
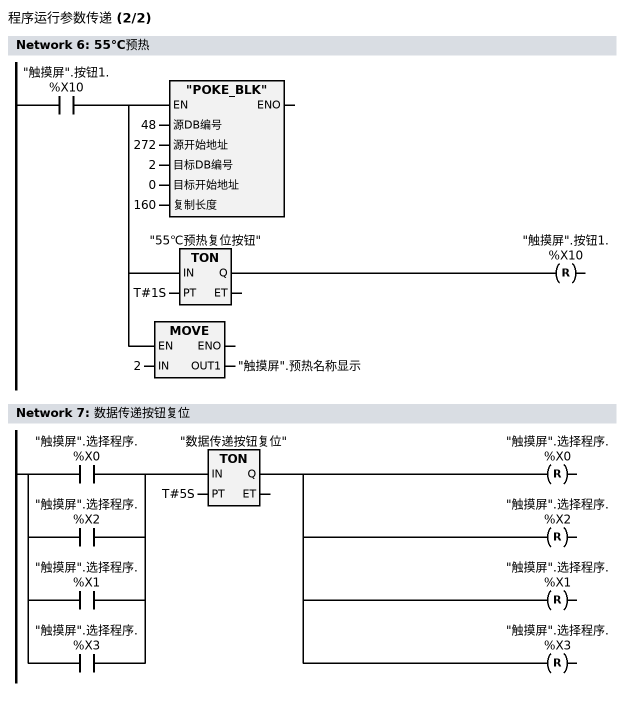
   #_w1 := "触摸屏".按钮1.%X10;
   IF #_w1 THEN "POKE_BLK"(源DB编号 := 48, 源开始地址 := 272, 目标DB编号 := 2, 目标开始地址 := 0, 复制长度 := 160); END_IF;
   "55℃预热复位按钮".TON(IN := #_w1, PT := T#1S);
   IF "55℃预热复位按钮".Q THEN "触摸屏".按钮1.%X10 := FALSE; END_IF;
   IF #_w1 THEN "触摸屏".预热名称显示 := 2; END_IF;
END_REGION

REGION Network 7: 数据传递按钮复位
   "数据传递按钮复位".TON(IN := "触摸屏".选择程序.%X0 OR "触摸屏".选择程序.%X2 OR "触摸屏".选择程序.%X1 OR "触摸屏".选择程序.%X3, PT := T#5S);
   IF "数据传递按钮复位".Q THEN
       "触摸屏".选择程序.%X0 := FALSE;
       "触摸屏".选择程序.%X2 := FALSE;
       "触摸屏".选择程序.%X1 := FALSE;
       "触摸屏".选择程序.%X3 := FALSE;
   END_IF;
END_REGION
END_FUNCTION_BLOCK

FUNCTION_BLOCK "程序数据编辑、保存（55℃参数除外）"   // FB22, LAD
{ S7_Optimized_Access := 'TRUE' }
VERSION : 0.1
   VAR
      沿1 : Bool;
      沿2 : Bool;
      沿3 : Bool;
      沿4 : Bool;
      沿5 : Bool;
      沿6 : Bool;
   END_VAR
   VAR_TEMP   // added for the SCL form of the ladder/FBD networks
      _w1 : Bool;
      _w2 : Bool;
      _w3 : Bool;
      _w4 : Bool;
      _w5 : Bool;
      _w6 : Bool;
      _w7 : Bool;
   END_VAR
BEGIN

REGION Network 1: 程序参数编辑选择
   // 1:37℃程序、2:药罐处理、3:泄露测试
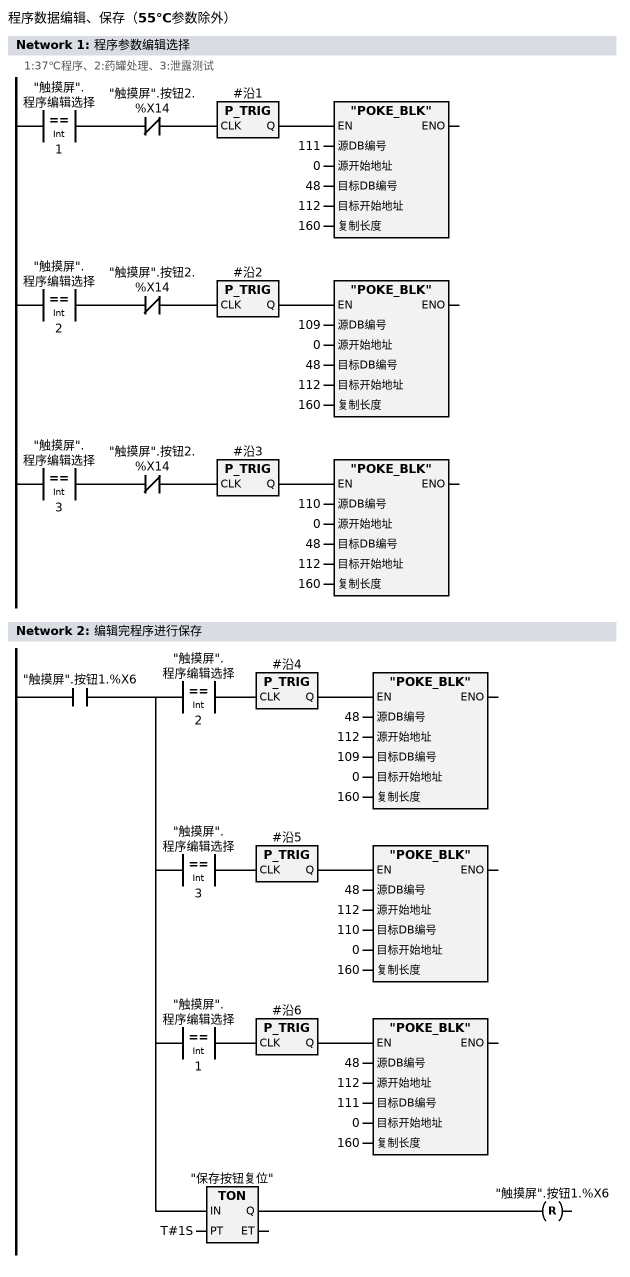
   RUNG wire#powerrail
      { S7_Templates := "SrcType := Int" } EQ_Contact(in1 := "触摸屏".程序编辑选择, in2 := 1)
      I_Contact( "触摸屏".按钮2.%X14 )
      P_Trig( #沿1 )
      "POKE_BLK"(源DB编号 := 111, 源开始地址 := 0, 目标DB编号 := 48, 目标开始地址 := 112, 复制长度 := 160)
   END_RUNG
   RUNG wire#powerrail
      { S7_Templates := "SrcType := Int" } EQ_Contact(in1 := "触摸屏".程序编辑选择, in2 := 2)
      I_Contact( "触摸屏".按钮2.%X14 )
      P_Trig( #沿2 )
      "POKE_BLK"(源DB编号 := 109, 源开始地址 := 0, 目标DB编号 := 48, 目标开始地址 := 112, 复制长度 := 160)
   END_RUNG
   RUNG wire#powerrail
      { S7_Templates := "SrcType := Int" } EQ_Contact(in1 := "触摸屏".程序编辑选择, in2 := 3)
      I_Contact( "触摸屏".按钮2.%X14 )
      P_Trig( #沿3 )
      "POKE_BLK"(源DB编号 := 110, 源开始地址 := 0, 目标DB编号 := 48, 目标开始地址 := 112, 复制长度 := 160)
   END_RUNG
   // the same network as SCL:
   #_w1 := ("触摸屏".程序编辑选择 = 1) AND NOT "触摸屏".按钮2.%X14;
   #_w2 := #_w1 AND NOT #沿1;   // rising edge
   #沿1 := #_w1;
   IF #_w2 THEN "POKE_BLK"(源DB编号 := 111, 源开始地址 := 0, 目标DB编号 := 48, 目标开始地址 := 112, 复制长度 := 160); END_IF;
   #_w3 := ("触摸屏".程序编辑选择 = 2) AND NOT "触摸屏".按钮2.%X14;
   #_w4 := #_w3 AND NOT #沿2;   // rising edge
   #沿2 := #_w3;
   IF #_w4 THEN "POKE_BLK"(源DB编号 := 109, 源开始地址 := 0, 目标DB编号 := 48, 目标开始地址 := 112, 复制长度 := 160); END_IF;
   #_w5 := ("触摸屏".程序编辑选择 = 3) AND NOT "触摸屏".按钮2.%X14;
   #_w6 := #_w5 AND NOT #沿3;   // rising edge
   #沿3 := #_w5;
   IF #_w6 THEN "POKE_BLK"(源DB编号 := 110, 源开始地址 := 0, 目标DB编号 := 48, 目标开始地址 := 112, 复制长度 := 160); END_IF;
END_REGION

REGION Network 2: 编辑完程序进行保存
   #_w1 := "触摸屏".按钮1.%X6 AND ("触摸屏".程序编辑选择 = 2);
   #_w2 := #_w1 AND NOT #沿4;   // rising edge
   #沿4 := #_w1;
   #_w3 := "触摸屏".按钮1.%X6;
   IF #_w2 THEN "POKE_BLK"(源DB编号 := 48, 源开始地址 := 112, 目标DB编号 := 109, 目标开始地址 := 0, 复制长度 := 160); END_IF;
   #_w4 := #_w3 AND ("触摸屏".程序编辑选择 = 3);
   #_w5 := #_w4 AND NOT #沿5;   // rising edge
   #沿5 := #_w4;
   IF #_w5 THEN "POKE_BLK"(源DB编号 := 48, 源开始地址 := 112, 目标DB编号 := 110, 目标开始地址 := 0, 复制长度 := 160); END_IF;
   #_w6 := #_w3 AND ("触摸屏".程序编辑选择 = 1);
   #_w7 := #_w6 AND NOT #沿6;   // rising edge
   #沿6 := #_w6;
   IF #_w7 THEN "POKE_BLK"(源DB编号 := 48, 源开始地址 := 112, 目标DB编号 := 111, 目标开始地址 := 0, 复制长度 := 160); END_IF;
   "保存按钮复位".TON(IN := #_w3, PT := T#1S);
   IF "保存按钮复位".Q THEN "触摸屏".按钮1.%X6 := FALSE; END_IF;
END_REGION
END_FUNCTION_BLOCK

FUNCTION "POKE_BLK" : Void   // FC2, SCL
{ S7_Optimized_Access := 'TRUE' }
VERSION : 0.1
   VAR_INPUT
      源DB编号 : Int;
      源开始地址 : Int;
      目标DB编号 : Int;
      目标开始地址 : Int;
      复制长度 : Int;
   END_VAR
BEGIN
   POKE_BLK(area_src:=16#84,
            dbNumber_src:=#源DB编号,
            byteOffset_src:=#源开始地址,
            area_dest:=16#84,
            dbNumber_dest:=#目标DB编号,
            byteOffset_dest:=#目标开始地址,
            count:=#复制长度);
END_FUNCTION

// folder: 8输入检测

FUNCTION "模拟量转换函数" : Void   // FC3, LAD
{ S7_Optimized_Access := 'TRUE' }
VERSION : 0.1
   VAR_INPUT
      模拟量输入最小值 : UInt;
      模拟量输入最大值 : UInt;
      模拟量输入值 : UInt;
      物理量最小值 : Real;
      物理量最大值 : Real;
      物理量校准值 : Int;
   END_VAR
   VAR_OUTPUT
      物理量输出值 : Int;
   END_VAR
   VAR_TEMP
      模拟量转换中间变量1 : Real;
      模拟量转换中间变量2 : Int;
      模拟量转换中间变量3 : Real;
      模拟量转换中间变量4 : UInt;
      模拟量转换最小值 : Int;
      模拟量转换最大值 : Int;
   END_VAR
BEGIN

REGION Network 1
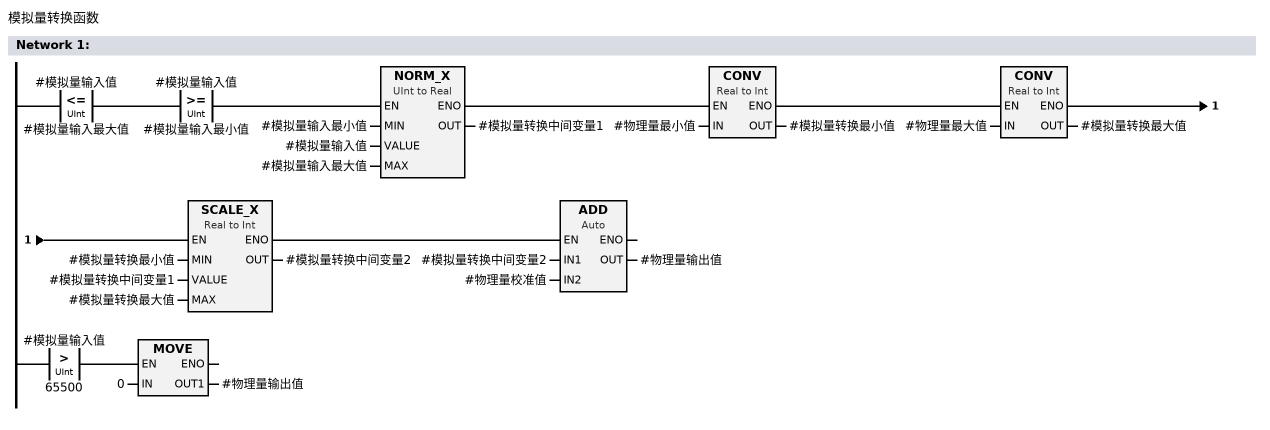
   RUNG wire#powerrail
      { S7_Templates := "SrcType := UInt" } LE_Contact(in1 := #模拟量输入值, in2 := #模拟量输入最大值)
      { S7_Templates := "SrcType := UInt" } GE_Contact(in1 := #模拟量输入值, in2 := #模拟量输入最小值)
      { S7_Templates := "[SrcType := UInt, DestType := Real]" } Normalize(min := #模拟量输入最小值, value := #模拟量输入值, max := #模拟量输入最大值, out => #模拟量转换中间变量1)
      { S7_Templates := "[SrcType := Real, DestType := Int]" } Convert(in := #物理量最小值, out => #模拟量转换最小值)
      { S7_Templates := "[SrcType := Real, DestType := Int]" } Convert(in := #物理量最大值, out => #模拟量转换最大值)
      { S7_Templates := "[SrcType := Real, DestType := Int]" } Scale(min := #模拟量转换最小值, value := #模拟量转换中间变量1, max := #模拟量转换最大值, out => #模拟量转换中间变量2)
      Add(in1 := #模拟量转换中间变量2, in2 := #物理量校准值, out => #物理量输出值)
   END_RUNG
   RUNG wire#powerrail
      { S7_Templates := "SrcType := UInt" } GT_Contact(in1 := #模拟量输入值, in2 := 65500)
      Move(in := 0, out1 => #物理量输出值)
   END_RUNG
   // the same network as SCL:
   IF (#模拟量输入值 <= #模拟量输入最大值) AND (#模拟量输入值 >= #模拟量输入最小值) THEN
       #模拟量转换中间变量1 := NORM_X(MIN := #模拟量输入最小值, VALUE := #模拟量输入值, MAX := #模拟量输入最大值);
       #模拟量转换最小值 := REAL_TO_INT(#物理量最小值);
       #模拟量转换最大值 := REAL_TO_INT(#物理量最大值);
       #模拟量转换中间变量2 := SCALE_X(MIN := #模拟量转换最小值, VALUE := #模拟量转换中间变量1, MAX := #模拟量转换最大值);
       #物理量输出值 := #模拟量转换中间变量2 + #物理量校准值;
   END_IF;
   IF #模拟量输入值 > 65500 THEN #物理量输出值 := 0; END_IF;
END_REGION
END_FUNCTION

FUNCTION "输入检测" : Void   // FC4, LAD
{ S7_Optimized_Access := 'TRUE' }
VERSION : 0.1
BEGIN

REGION Network 1: 数字量输入信号全部转到DI输入映像区
   // DI1.%X0：空压机保护
   // DI1.%X1：真空泵保护
   // DI1.%X2：前门电机过载
   // DI1.%X3：前门脚踢开关
   // DI1.%X4：后门脚踢开关
   // DI1.%X5：排气压力开关
   // DI1.%X6：关机确认信号
   // DI1.%X7：前门开位
   // DI1.%X8：前门关位
   // DI1.%X9：前门障碍
   // DI1.%X10：穿刺气缸位
   // DI1.%X11：水箱上水位
   // DI1.%X12：水箱下水位
   // DI1.%X13：压缩气压力检测
   // DI1.%X14：真空泵2保护
   // DI1.%X15：后门开位
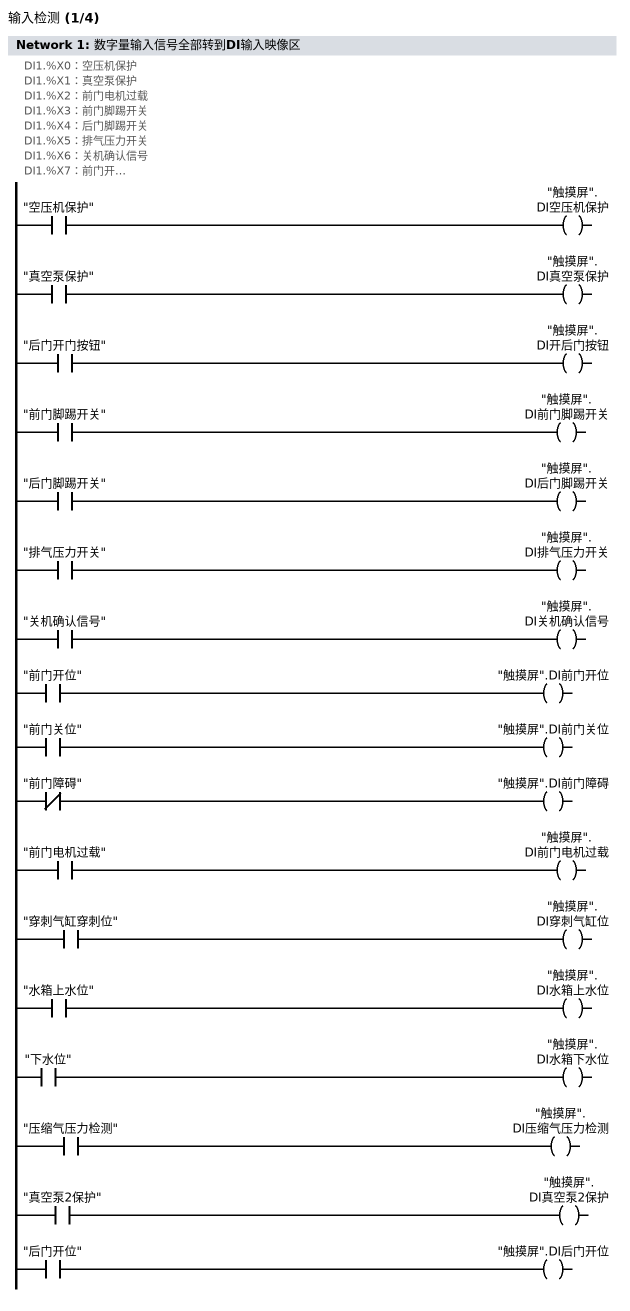
   RUNG wire#powerrail
      Contact( "空压机保护" )
      Coil( "触摸屏".DI空压机保护 )
   END_RUNG
   RUNG wire#powerrail
      Contact( "真空泵保护" )
      Coil( "触摸屏".DI真空泵保护 )
   END_RUNG
   RUNG wire#powerrail
      Contact( "后门开门按钮" )
      Coil( "触摸屏".DI开后门按钮 )
   END_RUNG
   RUNG wire#powerrail
      Contact( "前门脚踢开关" )
      Coil( "触摸屏".DI前门脚踢开关 )
   END_RUNG
   RUNG wire#powerrail
      Contact( "后门脚踢开关" )
      Coil( "触摸屏".DI后门脚踢开关 )
   END_RUNG
   RUNG wire#powerrail
      Contact( "排气压力开关" )
      Coil( "触摸屏".DI排气压力开关 )
   END_RUNG
   RUNG wire#powerrail
      Contact( "关机确认信号" )
      Coil( "触摸屏".DI关机确认信号 )
   END_RUNG
   RUNG wire#powerrail
      Contact( "前门开位" )
      Coil( "触摸屏".DI前门开位 )
   END_RUNG
   RUNG wire#powerrail
      Contact( "前门关位" )
      Coil( "触摸屏".DI前门关位 )
   END_RUNG
   RUNG wire#powerrail
      I_Contact( "前门障碍" )
      Coil( "触摸屏".DI前门障碍 )
   END_RUNG
   RUNG wire#powerrail
      Contact( "前门电机过载" )
      Coil( "触摸屏".DI前门电机过载 )
   END_RUNG
   RUNG wire#powerrail
      Contact( "穿刺气缸穿刺位" )
      Coil( "触摸屏".DI穿刺气缸位 )
   END_RUNG
   RUNG wire#powerrail
      Contact( "水箱上水位" )
      Coil( "触摸屏".DI水箱上水位 )
   END_RUNG
   RUNG wire#powerrail
      Contact( "下水位" )
      Coil( "触摸屏".DI水箱下水位 )
   END_RUNG
   RUNG wire#powerrail
      Contact( "压缩气压力检测" )
      Coil( "触摸屏".DI压缩气压力检测 )
   END_RUNG
   RUNG wire#powerrail
      Contact( "真空泵2保护" )
      Coil( "触摸屏".DI真空泵2保护 )
   END_RUNG
   RUNG wire#powerrail
      Contact( "后门开位" )
      Coil( "触摸屏".DI后门开位 )
   END_RUNG
   // the same network as SCL:
   "触摸屏".DI空压机保护 := "空压机保护";
   "触摸屏".DI真空泵保护 := "真空泵保护";
   "触摸屏".DI开后门按钮 := "后门开门按钮";
   "触摸屏".DI前门脚踢开关 := "前门脚踢开关";
   "触摸屏".DI后门脚踢开关 := "后门脚踢开关";
   "触摸屏".DI排气压力开关 := "排气压力开关";
   "触摸屏".DI关机确认信号 := "关机确认信号";
   "触摸屏".DI前门开位 := "前门开位";
   "触摸屏".DI前门关位 := "前门关位";
   "触摸屏".DI前门障碍 := NOT "前门障碍";
   "触摸屏".DI前门电机过载 := "前门电机过载";
   "触摸屏".DI穿刺气缸位 := "穿刺气缸穿刺位";
   "触摸屏".DI水箱上水位 := "水箱上水位";
   "触摸屏".DI水箱下水位 := "下水位";
   "触摸屏".DI压缩气压力检测 := "压缩气压力检测";
   "触摸屏".DI真空泵2保护 := "真空泵2保护";
   "触摸屏".DI后门开位 := "后门开位";
END_REGION

REGION Network 2
   // DI2.%X0：后门关位
   // DI2.%X1：后门障碍
   // DI2.%X2：急停按钮
   // DI2.%X3：后门电机过载
   // DI2.%X4：空压机过载保护
   // DI2.%X5：真空泵1过载
   // DI2.%X6：真空泵2过载
   // DI2.%X7：开后门按钮
   // DI2.%X8：关后门按钮
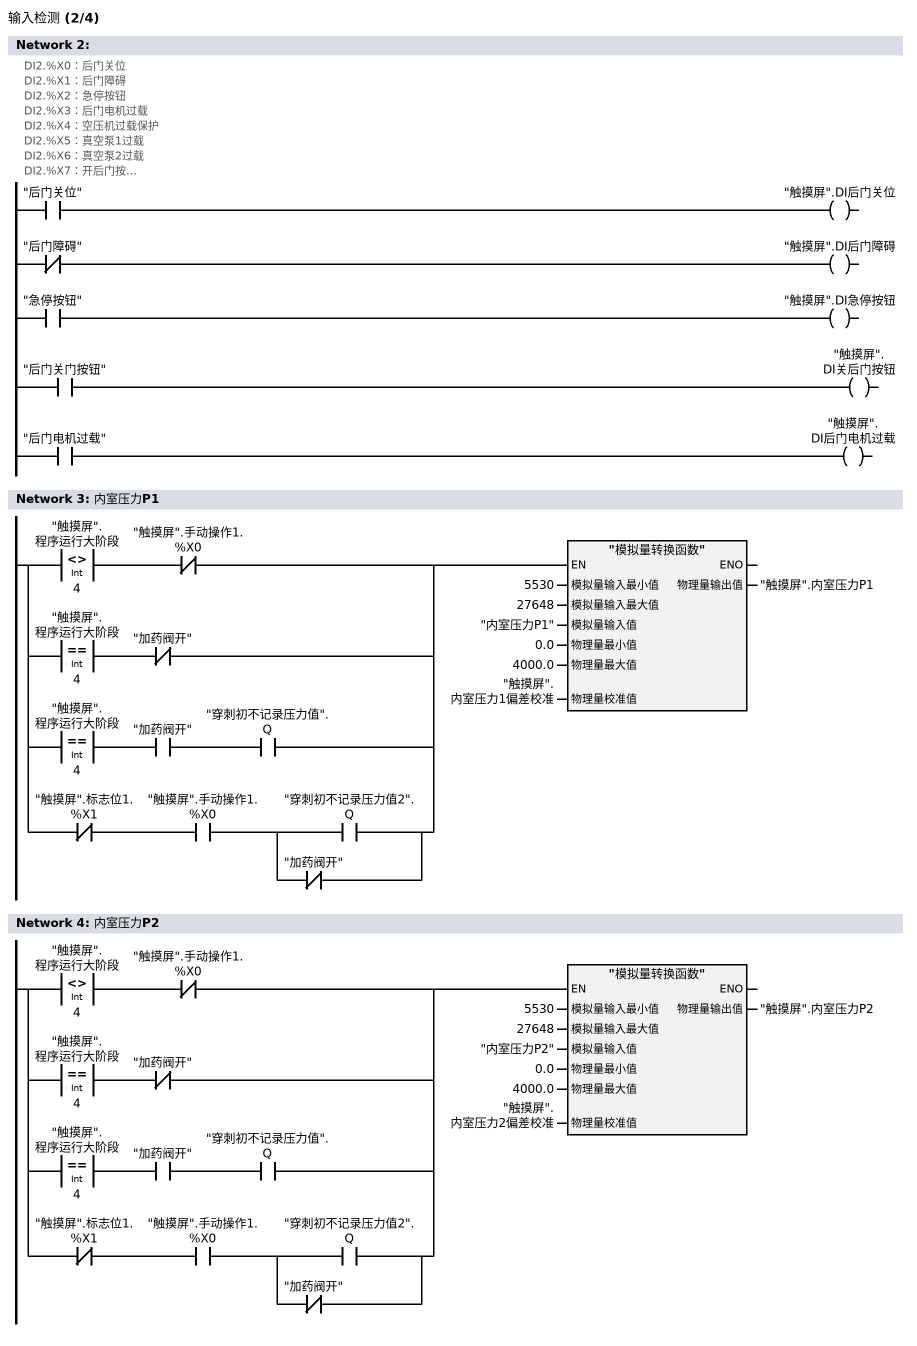
   RUNG wire#powerrail
      Contact( "后门关位" )
      Coil( "触摸屏".DI后门关位 )
   END_RUNG
   RUNG wire#powerrail
      I_Contact( "后门障碍" )
      Coil( "触摸屏".DI后门障碍 )
   END_RUNG
   RUNG wire#powerrail
      Contact( "急停按钮" )
      Coil( "触摸屏".DI急停按钮 )
   END_RUNG
   RUNG wire#powerrail
      Contact( "后门关门按钮" )
      Coil( "触摸屏".DI关后门按钮 )
   END_RUNG
   RUNG wire#powerrail
      Contact( "后门电机过载" )
      Coil( "触摸屏".DI后门电机过载 )
   END_RUNG
   // the same network as SCL:
   "触摸屏".DI后门关位 := "后门关位";
   "触摸屏".DI后门障碍 := NOT "后门障碍";
   "触摸屏".DI急停按钮 := "急停按钮";
   "触摸屏".DI关后门按钮 := "后门关门按钮";
   "触摸屏".DI后门电机过载 := "后门电机过载";
END_REGION

REGION Network 3: 内室压力P1
   RUNG wire#powerrail
      { S7_Templates := "SrcType := Int" } NE_Contact(in1 := "触摸屏".程序运行大阶段, in2 := 4)
      I_Contact( "触摸屏".手动操作1.%X0 )
      wire#w1
      "模拟量转换函数"(模拟量输入最小值 := 5530, 模拟量输入最大值 := 27648, 模拟量输入值 := "内室压力P1", 物理量最小值 := 0.0, 物理量最大值 := 4000.0, 物理量校准值 := "触摸屏".内室压力1偏差校准, 物理量输出值 => "触摸屏".内室压力P1)
   END_RUNG
   RUNG wire#powerrail
      { S7_Templates := "SrcType := Int" } EQ_Contact(in1 := "触摸屏".程序运行大阶段, in2 := 4)
      I_Contact( "加药阀开" )
   END_RUNG wire#w1
   RUNG wire#powerrail
      { S7_Templates := "SrcType := Int" } EQ_Contact(in1 := "触摸屏".程序运行大阶段, in2 := 4)
      Contact( "加药阀开" )
      Contact( "穿刺初不记录压力值".Q )
   END_RUNG wire#w1
   RUNG wire#powerrail
      I_Contact( "触摸屏".标志位1.%X1 )
      Contact( "触摸屏".手动操作1.%X0 )
      wire#w2
      Contact( "穿刺初不记录压力值2".Q )
   END_RUNG wire#w1
   RUNG wire#w2
      I_Contact( "加药阀开" )
   END_RUNG wire#w1
   // the same network as SCL:
   IF (("触摸屏".程序运行大阶段 <> 4) AND NOT "触摸屏".手动操作1.%X0) OR (("触摸屏".程序运行大阶段 = 4) AND NOT "加药阀开") OR (("触摸屏".程序运行大阶段 = 4) AND "加药阀开" AND "穿刺初不记录压力值".Q) OR (NOT "触摸屏".标志位1.%X1 AND "触摸屏".手动操作1.%X0 AND ("穿刺初不记录压力值2".Q OR NOT "加药阀开")) THEN
       "模拟量转换函数"(模拟量输入最小值 := 5530,
                 模拟量输入最大值 := 27648,
                 模拟量输入值 := "内室压力P1",
                 物理量最小值 := 0.0,
                 物理量最大值 := 4000.0,
                 物理量校准值 := "触摸屏".内室压力1偏差校准,
                 物理量输出值 => "触摸屏".内室压力P1);
   END_IF;
END_REGION

REGION Network 4: 内室压力P2
   RUNG wire#powerrail
      { S7_Templates := "SrcType := Int" } NE_Contact(in1 := "触摸屏".程序运行大阶段, in2 := 4)
      I_Contact( "触摸屏".手动操作1.%X0 )
      wire#w1
      "模拟量转换函数"(模拟量输入最小值 := 5530, 模拟量输入最大值 := 27648, 模拟量输入值 := "内室压力P2", 物理量最小值 := 0.0, 物理量最大值 := 4000.0, 物理量校准值 := "触摸屏".内室压力2偏差校准, 物理量输出值 => "触摸屏".内室压力P2)
   END_RUNG
   RUNG wire#powerrail
      { S7_Templates := "SrcType := Int" } EQ_Contact(in1 := "触摸屏".程序运行大阶段, in2 := 4)
      I_Contact( "加药阀开" )
   END_RUNG wire#w1
   RUNG wire#powerrail
      { S7_Templates := "SrcType := Int" } EQ_Contact(in1 := "触摸屏".程序运行大阶段, in2 := 4)
      Contact( "加药阀开" )
      Contact( "穿刺初不记录压力值".Q )
   END_RUNG wire#w1
   RUNG wire#powerrail
      I_Contact( "触摸屏".标志位1.%X1 )
      Contact( "触摸屏".手动操作1.%X0 )
      wire#w2
      Contact( "穿刺初不记录压力值2".Q )
   END_RUNG wire#w1
   RUNG wire#w2
      I_Contact( "加药阀开" )
   END_RUNG wire#w1
   // the same network as SCL:
   IF (("触摸屏".程序运行大阶段 <> 4) AND NOT "触摸屏".手动操作1.%X0) OR (("触摸屏".程序运行大阶段 = 4) AND NOT "加药阀开") OR (("触摸屏".程序运行大阶段 = 4) AND "加药阀开" AND "穿刺初不记录压力值".Q) OR (NOT "触摸屏".标志位1.%X1 AND "触摸屏".手动操作1.%X0 AND ("穿刺初不记录压力值2".Q OR NOT "加药阀开")) THEN
       "模拟量转换函数"(模拟量输入最小值 := 5530,
                 模拟量输入最大值 := 27648,
                 模拟量输入值 := "内室压力P2",
                 物理量最小值 := 0.0,
                 物理量最大值 := 4000.0,
                 物理量校准值 := "触摸屏".内室压力2偏差校准,
                 物理量输出值 => "触摸屏".内室压力P2);
   END_IF;
END_REGION

REGION Network 5: 内室温度T1
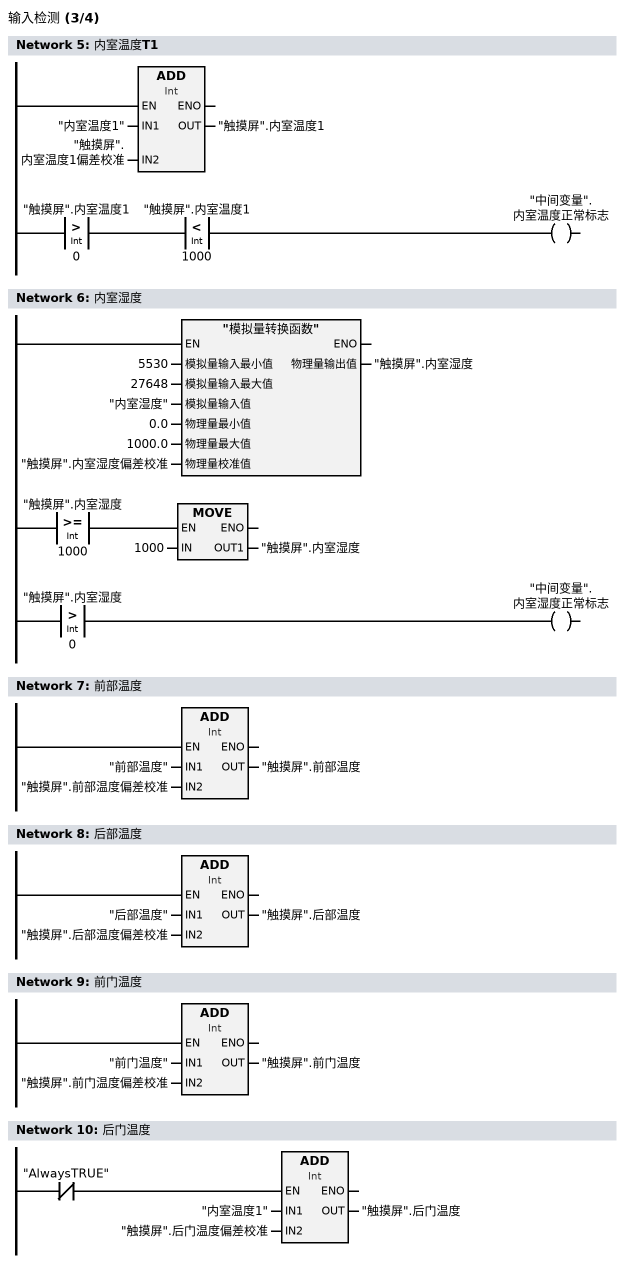
   RUNG wire#powerrail
      { S7_Templates := "SrcType := Int" } Add(in1 := "内室温度1", in2 := "触摸屏".内室温度1偏差校准, out => "触摸屏".内室温度1)
   END_RUNG
   RUNG wire#powerrail
      { S7_Templates := "SrcType := Int" } GT_Contact(in1 := "触摸屏".内室温度1, in2 := 0)
      { S7_Templates := "SrcType := Int" } LT_Contact(in1 := "触摸屏".内室温度1, in2 := 1000)
      Coil( "中间变量".内室温度正常标志 )
   END_RUNG
   // the same network as SCL:
   "触摸屏".内室温度1 := "内室温度1" + "触摸屏".内室温度1偏差校准;
   "中间变量".内室温度正常标志 := ("触摸屏".内室温度1 > 0) AND ("触摸屏".内室温度1 < 1000);
END_REGION

REGION Network 6: 内室湿度
   RUNG wire#powerrail
      "模拟量转换函数"(模拟量输入最小值 := 5530, 模拟量输入最大值 := 27648, 模拟量输入值 := "内室湿度", 物理量最小值 := 0.0, 物理量最大值 := 1000.0, 物理量校准值 := "触摸屏".内室湿度偏差校准, 物理量输出值 => "触摸屏".内室湿度)
   END_RUNG
   RUNG wire#powerrail
      { S7_Templates := "SrcType := Int" } GE_Contact(in1 := "触摸屏".内室湿度, in2 := 1000)
      Move(in := 1000, out1 => "触摸屏".内室湿度)
   END_RUNG
   RUNG wire#powerrail
      { S7_Templates := "SrcType := Int" } GT_Contact(in1 := "触摸屏".内室湿度, in2 := 0)
      Coil( "中间变量".内室湿度正常标志 )
   END_RUNG
   // the same network as SCL:
   "模拟量转换函数"(模拟量输入最小值 := 5530,
             模拟量输入最大值 := 27648,
             模拟量输入值 := "内室湿度",
             物理量最小值 := 0.0,
             物理量最大值 := 1000.0,
             物理量校准值 := "触摸屏".内室湿度偏差校准,
             物理量输出值 => "触摸屏".内室湿度);
   IF "触摸屏".内室湿度 >= 1000 THEN "触摸屏".内室湿度 := 1000; END_IF;
   "中间变量".内室湿度正常标志 := "触摸屏".内室湿度 > 0;
END_REGION

REGION Network 7: 前部温度
   RUNG wire#powerrail
      { S7_Templates := "SrcType := Int" } Add(in1 := "前部温度", in2 := "触摸屏".前部温度偏差校准, out => "触摸屏".前部温度)
   END_RUNG
   // the same network as SCL:
   "触摸屏".前部温度 := "前部温度" + "触摸屏".前部温度偏差校准;
END_REGION

REGION Network 8: 后部温度
   RUNG wire#powerrail
      { S7_Templates := "SrcType := Int" } Add(in1 := "后部温度", in2 := "触摸屏".后部温度偏差校准, out => "触摸屏".后部温度)
   END_RUNG
   // the same network as SCL:
   "触摸屏".后部温度 := "后部温度" + "触摸屏".后部温度偏差校准;
END_REGION

REGION Network 9: 前门温度
   RUNG wire#powerrail
      { S7_Templates := "SrcType := Int" } Add(in1 := "前门温度", in2 := "触摸屏".前门温度偏差校准, out => "触摸屏".前门温度)
   END_RUNG
   // the same network as SCL:
   "触摸屏".前门温度 := "前门温度" + "触摸屏".前门温度偏差校准;
END_REGION

REGION Network 10: 后门温度
   RUNG wire#powerrail
      I_Contact( "AlwaysTRUE" )
      { S7_Templates := "SrcType := Int" } Add(in1 := "内室温度1", in2 := "触摸屏".后门温度偏差校准, out => "触摸屏".后门温度)
   END_RUNG
   // the same network as SCL:
   IF NOT "AlwaysTRUE" THEN "触摸屏".后门温度 := "内室温度1" + "触摸屏".后门温度偏差校准; END_IF;
END_REGION

REGION Network 11: 汽化室温度
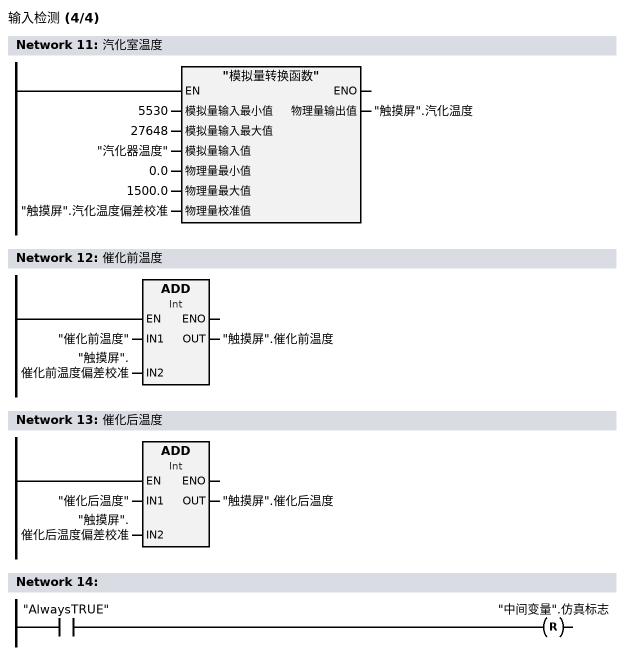
   RUNG wire#powerrail
      "模拟量转换函数"(模拟量输入最小值 := 5530, 模拟量输入最大值 := 27648, 模拟量输入值 := "汽化器温度", 物理量最小值 := 0.0, 物理量最大值 := 1500.0, 物理量校准值 := "触摸屏".汽化温度偏差校准, 物理量输出值 => "触摸屏".汽化温度)
   END_RUNG
   // the same network as SCL:
   "模拟量转换函数"(模拟量输入最小值 := 5530,
             模拟量输入最大值 := 27648,
             模拟量输入值 := "汽化器温度",
             物理量最小值 := 0.0,
             物理量最大值 := 1500.0,
             物理量校准值 := "触摸屏".汽化温度偏差校准,
             物理量输出值 => "触摸屏".汽化温度);
END_REGION

REGION Network 12: 催化前温度
   RUNG wire#powerrail
      { S7_Templates := "SrcType := Int" } Add(in1 := "催化前温度", in2 := "触摸屏".催化前温度偏差校准, out => "触摸屏".催化前温度)
   END_RUNG
   // the same network as SCL:
   "触摸屏".催化前温度 := "催化前温度" + "触摸屏".催化前温度偏差校准;
END_REGION

REGION Network 13: 催化后温度
   RUNG wire#powerrail
      { S7_Templates := "SrcType := Int" } Add(in1 := "催化后温度", in2 := "触摸屏".催化后温度偏差校准, out => "触摸屏".催化后温度)
   END_RUNG
   // the same network as SCL:
   "触摸屏".催化后温度 := "催化后温度" + "触摸屏".催化后温度偏差校准;
END_REGION

REGION Network 14
   RUNG wire#powerrail
      Contact( "AlwaysTRUE" )
      R_Coil( "中间变量".仿真标志 )
   END_RUNG
   // the same network as SCL:
   IF "AlwaysTRUE" THEN "中间变量".仿真标志 := FALSE; END_IF;
END_REGION
END_FUNCTION

FUNCTION "仿真输入检测" : Void   // FC8, LAD
{ S7_Optimized_Access := 'TRUE' }
VERSION : 0.1
   VAR_TEMP   // added for the SCL form of the ladder/FBD networks
      _w1 : Bool;
      _w2 : Bool;
      _w3 : Bool;
      _w4 : Bool;
   END_VAR
BEGIN

REGION Network 1: 数字量输入信号全部转到DI输入映像区
   // DI1.%X0：空压机保护
   // DI1.%X1：真空泵保护
   // DI1.%X2：前门电机过载
   // DI1.%X3：前门脚踢开关
   // DI1.%X4：后门脚踢开关
   // DI1.%X5：排气压力开关
   // DI1.%X6：关机确认信号
   // DI1.%X7：前门开位
   // DI1.%X8：前门关位
   // DI1.%X9：前门障碍
   // DI1.%X10：穿刺气缸位
   // DI1.%X11：水箱上水位
   // DI1.%X12：水箱下水位
   // DI1.%X13：压缩气压力检测
   // DI1.%X14：真空泵2保护
   // DI1.%X15：后门开位
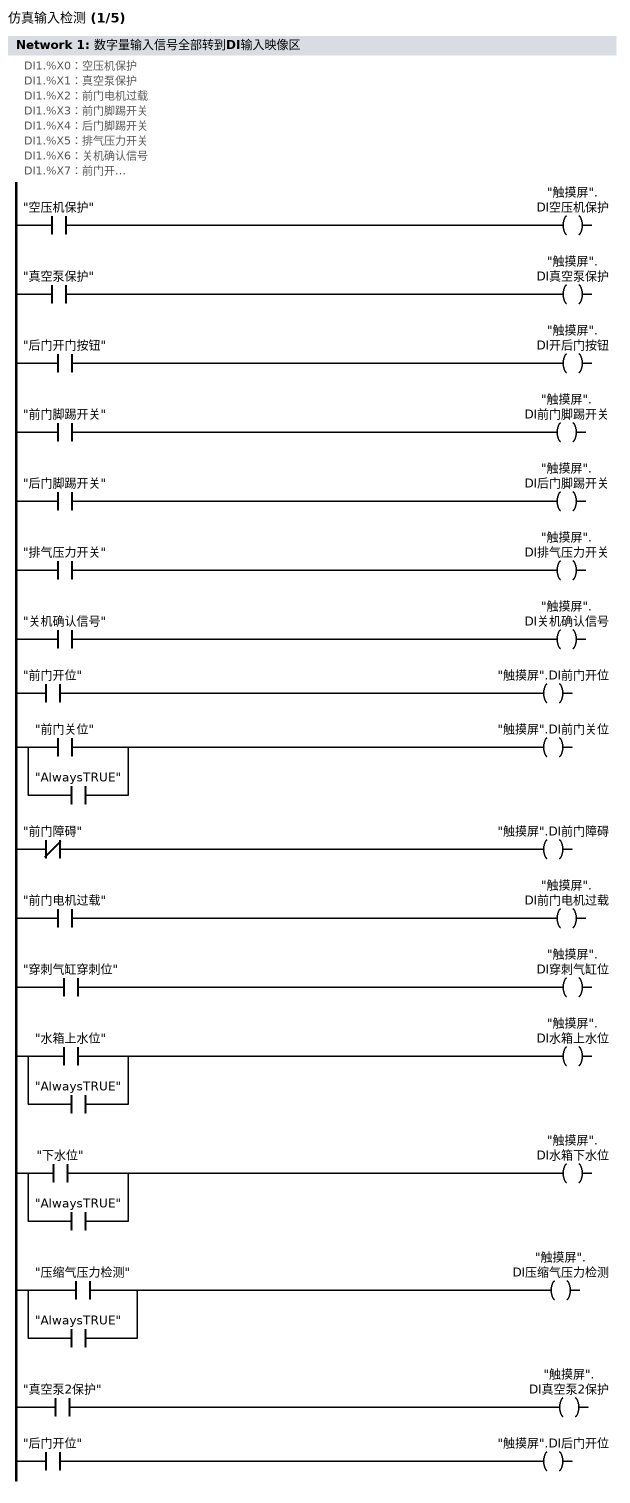
   RUNG wire#powerrail
      Contact( "空压机保护" )
      Coil( "触摸屏".DI空压机保护 )
   END_RUNG
   RUNG wire#powerrail
      Contact( "真空泵保护" )
      Coil( "触摸屏".DI真空泵保护 )
   END_RUNG
   RUNG wire#powerrail
      Contact( "后门开门按钮" )
      Coil( "触摸屏".DI开后门按钮 )
   END_RUNG
   RUNG wire#powerrail
      Contact( "前门脚踢开关" )
      Coil( "触摸屏".DI前门脚踢开关 )
   END_RUNG
   RUNG wire#powerrail
      Contact( "后门脚踢开关" )
      Coil( "触摸屏".DI后门脚踢开关 )
   END_RUNG
   RUNG wire#powerrail
      Contact( "排气压力开关" )
      Coil( "触摸屏".DI排气压力开关 )
   END_RUNG
   RUNG wire#powerrail
      Contact( "关机确认信号" )
      Coil( "触摸屏".DI关机确认信号 )
   END_RUNG
   RUNG wire#powerrail
      Contact( "前门开位" )
      Coil( "触摸屏".DI前门开位 )
   END_RUNG
   RUNG wire#powerrail
      Contact( "前门关位" )
      wire#w1
      Coil( "触摸屏".DI前门关位 )
   END_RUNG
   RUNG wire#powerrail
      Contact( "AlwaysTRUE" )
   END_RUNG wire#w1
   RUNG wire#powerrail
      I_Contact( "前门障碍" )
      Coil( "触摸屏".DI前门障碍 )
   END_RUNG
   RUNG wire#powerrail
      Contact( "前门电机过载" )
      Coil( "触摸屏".DI前门电机过载 )
   END_RUNG
   RUNG wire#powerrail
      Contact( "穿刺气缸穿刺位" )
      Coil( "触摸屏".DI穿刺气缸位 )
   END_RUNG
   RUNG wire#powerrail
      Contact( "水箱上水位" )
      wire#w2
      Coil( "触摸屏".DI水箱上水位 )
   END_RUNG
   RUNG wire#powerrail
      Contact( "AlwaysTRUE" )
   END_RUNG wire#w2
   RUNG wire#powerrail
      Contact( "下水位" )
      wire#w3
      Coil( "触摸屏".DI水箱下水位 )
   END_RUNG
   RUNG wire#powerrail
      Contact( "AlwaysTRUE" )
   END_RUNG wire#w3
   RUNG wire#powerrail
      Contact( "压缩气压力检测" )
      wire#w4
      Coil( "触摸屏".DI压缩气压力检测 )
   END_RUNG
   RUNG wire#powerrail
      Contact( "AlwaysTRUE" )
   END_RUNG wire#w4
   RUNG wire#powerrail
      Contact( "真空泵2保护" )
      Coil( "触摸屏".DI真空泵2保护 )
   END_RUNG
   RUNG wire#powerrail
      Contact( "后门开位" )
      Coil( "触摸屏".DI后门开位 )
   END_RUNG
   // the same network as SCL:
   "触摸屏".DI空压机保护 := "空压机保护";
   "触摸屏".DI真空泵保护 := "真空泵保护";
   "触摸屏".DI开后门按钮 := "后门开门按钮";
   "触摸屏".DI前门脚踢开关 := "前门脚踢开关";
   "触摸屏".DI后门脚踢开关 := "后门脚踢开关";
   "触摸屏".DI排气压力开关 := "排气压力开关";
   "触摸屏".DI关机确认信号 := "关机确认信号";
   "触摸屏".DI前门开位 := "前门开位";
   "触摸屏".DI前门关位 := "前门关位" OR "AlwaysTRUE";
   "触摸屏".DI前门障碍 := NOT "前门障碍";
   "触摸屏".DI前门电机过载 := "前门电机过载";
   "触摸屏".DI穿刺气缸位 := "穿刺气缸穿刺位";
   "触摸屏".DI水箱上水位 := "水箱上水位" OR "AlwaysTRUE";
   "触摸屏".DI水箱下水位 := "下水位" OR "AlwaysTRUE";
   "触摸屏".DI压缩气压力检测 := "压缩气压力检测" OR "AlwaysTRUE";
   "触摸屏".DI真空泵2保护 := "真空泵2保护";
   "触摸屏".DI后门开位 := "后门开位";
END_REGION

REGION Network 2
   // DI2.%X0：后门关位
   // DI2.%X1：后门障碍
   // DI2.%X2：急停按钮
   // DI2.%X3：后门电机过载
   // DI2.%X4：空压机过载保护
   // DI2.%X5：真空泵1过载
   // DI2.%X6：真空泵2过载
   // DI2.%X7：开后门按钮
   // DI2.%X8：关后门按钮
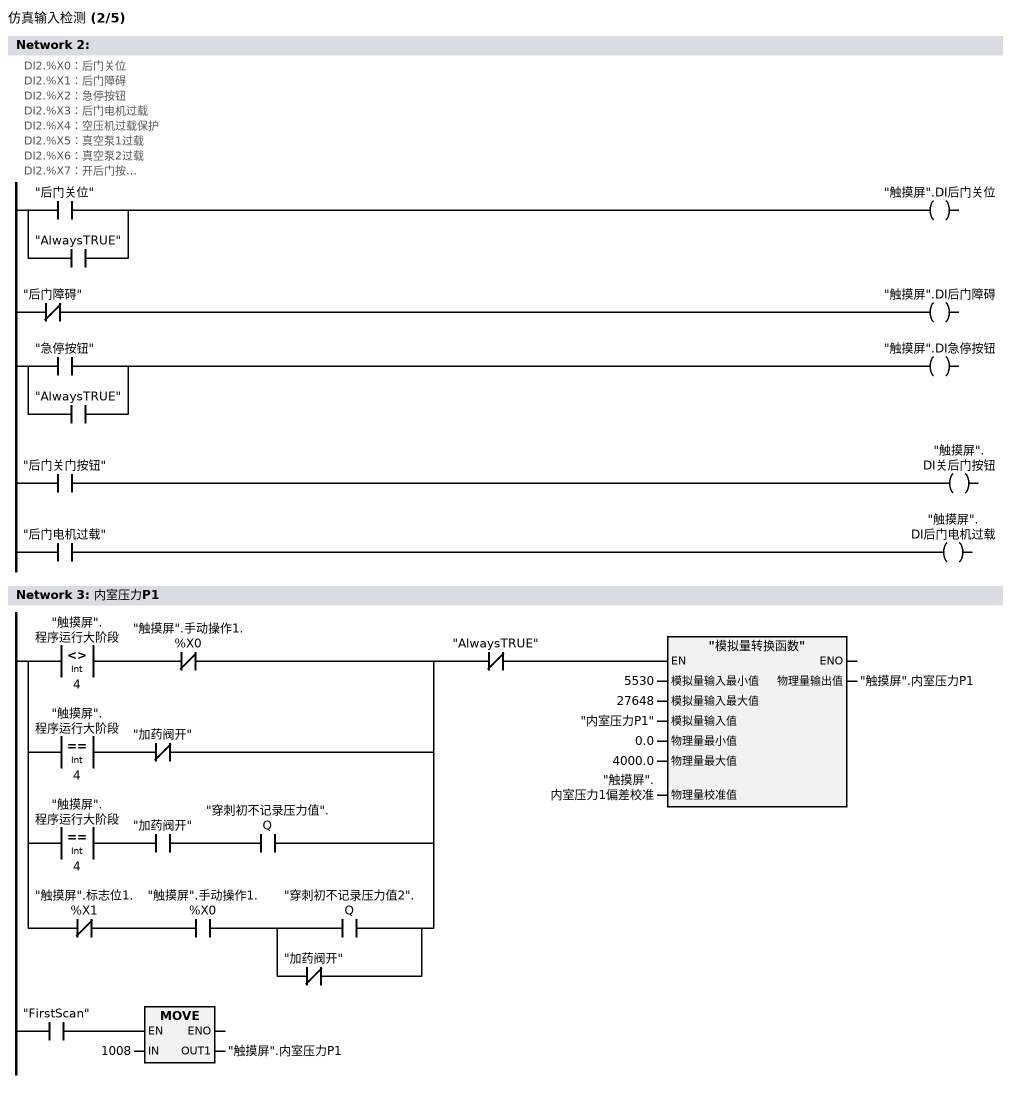
   RUNG wire#powerrail
      Contact( "后门关位" )
      wire#w1
      Coil( "触摸屏".DI后门关位 )
   END_RUNG
   RUNG wire#powerrail
      Contact( "AlwaysTRUE" )
   END_RUNG wire#w1
   RUNG wire#powerrail
      I_Contact( "后门障碍" )
      Coil( "触摸屏".DI后门障碍 )
   END_RUNG
   RUNG wire#powerrail
      Contact( "急停按钮" )
      wire#w2
      Coil( "触摸屏".DI急停按钮 )
   END_RUNG
   RUNG wire#powerrail
      Contact( "AlwaysTRUE" )
   END_RUNG wire#w2
   RUNG wire#powerrail
      Contact( "后门关门按钮" )
      Coil( "触摸屏".DI关后门按钮 )
   END_RUNG
   RUNG wire#powerrail
      Contact( "后门电机过载" )
      Coil( "触摸屏".DI后门电机过载 )
   END_RUNG
   // the same network as SCL:
   "触摸屏".DI后门关位 := "后门关位" OR "AlwaysTRUE";
   "触摸屏".DI后门障碍 := NOT "后门障碍";
   "触摸屏".DI急停按钮 := "急停按钮" OR "AlwaysTRUE";
   "触摸屏".DI关后门按钮 := "后门关门按钮";
   "触摸屏".DI后门电机过载 := "后门电机过载";
END_REGION

REGION Network 3: 内室压力P1
   RUNG wire#powerrail
      { S7_Templates := "SrcType := Int" } NE_Contact(in1 := "触摸屏".程序运行大阶段, in2 := 4)
      I_Contact( "触摸屏".手动操作1.%X0 )
      wire#w1
      I_Contact( "AlwaysTRUE" )
      "模拟量转换函数"(模拟量输入最小值 := 5530, 模拟量输入最大值 := 27648, 模拟量输入值 := "内室压力P1", 物理量最小值 := 0.0, 物理量最大值 := 4000.0, 物理量校准值 := "触摸屏".内室压力1偏差校准, 物理量输出值 => "触摸屏".内室压力P1)
   END_RUNG
   RUNG wire#powerrail
      { S7_Templates := "SrcType := Int" } EQ_Contact(in1 := "触摸屏".程序运行大阶段, in2 := 4)
      I_Contact( "加药阀开" )
   END_RUNG wire#w1
   RUNG wire#powerrail
      { S7_Templates := "SrcType := Int" } EQ_Contact(in1 := "触摸屏".程序运行大阶段, in2 := 4)
      Contact( "加药阀开" )
      Contact( "穿刺初不记录压力值".Q )
   END_RUNG wire#w1
   RUNG wire#powerrail
      I_Contact( "触摸屏".标志位1.%X1 )
      Contact( "触摸屏".手动操作1.%X0 )
      wire#w2
      Contact( "穿刺初不记录压力值2".Q )
   END_RUNG wire#w1
   RUNG wire#w2
      I_Contact( "加药阀开" )
   END_RUNG wire#w1
   RUNG wire#powerrail
      Contact( "FirstScan" )
      Move(in := 1008, out1 => "触摸屏".内室压力P1)
   END_RUNG
   // the same network as SCL:
   IF ((("触摸屏".程序运行大阶段 <> 4) AND NOT "触摸屏".手动操作1.%X0) OR (("触摸屏".程序运行大阶段 = 4) AND NOT "加药阀开") OR (("触摸屏".程序运行大阶段 = 4) AND "加药阀开" AND "穿刺初不记录压力值".Q) OR (NOT "触摸屏".标志位1.%X1 AND "触摸屏".手动操作1.%X0 AND ("穿刺初不记录压力值2".Q OR NOT "加药阀开"))) AND NOT "AlwaysTRUE" THEN
       "模拟量转换函数"(模拟量输入最小值 := 5530,
                 模拟量输入最大值 := 27648,
                 模拟量输入值 := "内室压力P1",
                 物理量最小值 := 0.0,
                 物理量最大值 := 4000.0,
                 物理量校准值 := "触摸屏".内室压力1偏差校准,
                 物理量输出值 => "触摸屏".内室压力P1);
   END_IF;
   IF "FirstScan" THEN "触摸屏".内室压力P1 := 1008; END_IF;
END_REGION

REGION Network 4: 内室压力P2
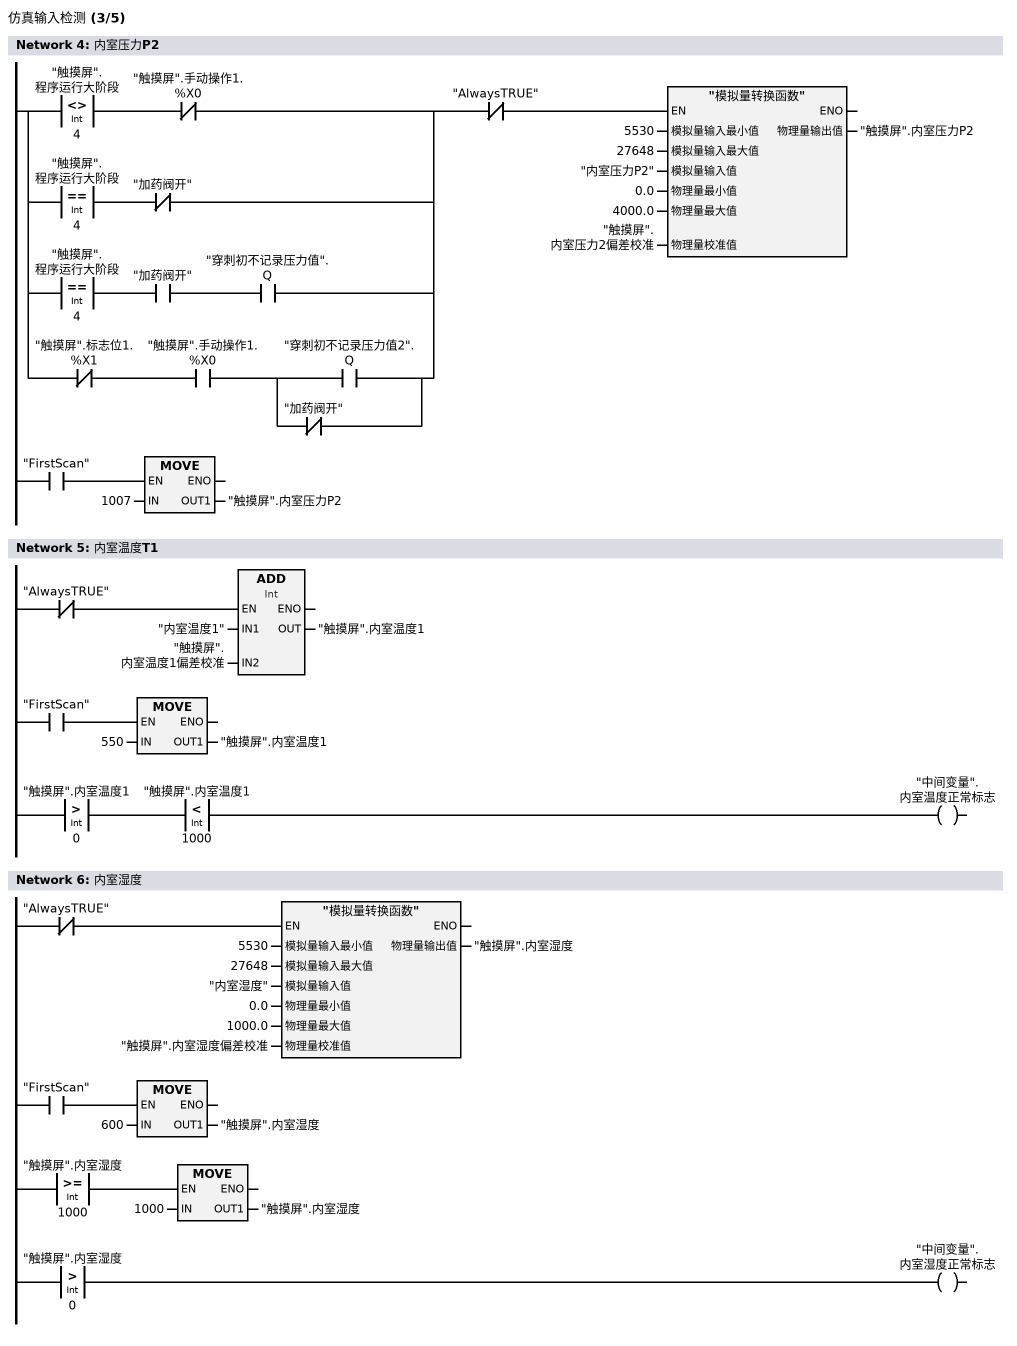
   RUNG wire#powerrail
      { S7_Templates := "SrcType := Int" } NE_Contact(in1 := "触摸屏".程序运行大阶段, in2 := 4)
      I_Contact( "触摸屏".手动操作1.%X0 )
      wire#w1
      I_Contact( "AlwaysTRUE" )
      "模拟量转换函数"(模拟量输入最小值 := 5530, 模拟量输入最大值 := 27648, 模拟量输入值 := "内室压力P2", 物理量最小值 := 0.0, 物理量最大值 := 4000.0, 物理量校准值 := "触摸屏".内室压力2偏差校准, 物理量输出值 => "触摸屏".内室压力P2)
   END_RUNG
   RUNG wire#powerrail
      { S7_Templates := "SrcType := Int" } EQ_Contact(in1 := "触摸屏".程序运行大阶段, in2 := 4)
      I_Contact( "加药阀开" )
   END_RUNG wire#w1
   RUNG wire#powerrail
      { S7_Templates := "SrcType := Int" } EQ_Contact(in1 := "触摸屏".程序运行大阶段, in2 := 4)
      Contact( "加药阀开" )
      Contact( "穿刺初不记录压力值".Q )
   END_RUNG wire#w1
   RUNG wire#powerrail
      I_Contact( "触摸屏".标志位1.%X1 )
      Contact( "触摸屏".手动操作1.%X0 )
      wire#w2
      Contact( "穿刺初不记录压力值2".Q )
   END_RUNG wire#w1
   RUNG wire#w2
      I_Contact( "加药阀开" )
   END_RUNG wire#w1
   RUNG wire#powerrail
      Contact( "FirstScan" )
      Move(in := 1007, out1 => "触摸屏".内室压力P2)
   END_RUNG
   // the same network as SCL:
   IF ((("触摸屏".程序运行大阶段 <> 4) AND NOT "触摸屏".手动操作1.%X0) OR (("触摸屏".程序运行大阶段 = 4) AND NOT "加药阀开") OR (("触摸屏".程序运行大阶段 = 4) AND "加药阀开" AND "穿刺初不记录压力值".Q) OR (NOT "触摸屏".标志位1.%X1 AND "触摸屏".手动操作1.%X0 AND ("穿刺初不记录压力值2".Q OR NOT "加药阀开"))) AND NOT "AlwaysTRUE" THEN
       "模拟量转换函数"(模拟量输入最小值 := 5530,
                 模拟量输入最大值 := 27648,
                 模拟量输入值 := "内室压力P2",
                 物理量最小值 := 0.0,
                 物理量最大值 := 4000.0,
                 物理量校准值 := "触摸屏".内室压力2偏差校准,
                 物理量输出值 => "触摸屏".内室压力P2);
   END_IF;
   IF "FirstScan" THEN "触摸屏".内室压力P2 := 1007; END_IF;
END_REGION

REGION Network 5: 内室温度T1
   RUNG wire#powerrail
      I_Contact( "AlwaysTRUE" )
      { S7_Templates := "SrcType := Int" } Add(in1 := "内室温度1", in2 := "触摸屏".内室温度1偏差校准, out => "触摸屏".内室温度1)
   END_RUNG
   RUNG wire#powerrail
      Contact( "FirstScan" )
      Move(in := 550, out1 => "触摸屏".内室温度1)
   END_RUNG
   RUNG wire#powerrail
      { S7_Templates := "SrcType := Int" } GT_Contact(in1 := "触摸屏".内室温度1, in2 := 0)
      { S7_Templates := "SrcType := Int" } LT_Contact(in1 := "触摸屏".内室温度1, in2 := 1000)
      Coil( "中间变量".内室温度正常标志 )
   END_RUNG
   // the same network as SCL:
   IF NOT "AlwaysTRUE" THEN "触摸屏".内室温度1 := "内室温度1" + "触摸屏".内室温度1偏差校准; END_IF;
   IF "FirstScan" THEN "触摸屏".内室温度1 := 550; END_IF;
   "中间变量".内室温度正常标志 := ("触摸屏".内室温度1 > 0) AND ("触摸屏".内室温度1 < 1000);
END_REGION

REGION Network 6: 内室湿度
   RUNG wire#powerrail
      I_Contact( "AlwaysTRUE" )
      "模拟量转换函数"(模拟量输入最小值 := 5530, 模拟量输入最大值 := 27648, 模拟量输入值 := "内室湿度", 物理量最小值 := 0.0, 物理量最大值 := 1000.0, 物理量校准值 := "触摸屏".内室湿度偏差校准, 物理量输出值 => "触摸屏".内室湿度)
   END_RUNG
   RUNG wire#powerrail
      Contact( "FirstScan" )
      Move(in := 600, out1 => "触摸屏".内室湿度)
   END_RUNG
   RUNG wire#powerrail
      { S7_Templates := "SrcType := Int" } GE_Contact(in1 := "触摸屏".内室湿度, in2 := 1000)
      Move(in := 1000, out1 => "触摸屏".内室湿度)
   END_RUNG
   RUNG wire#powerrail
      { S7_Templates := "SrcType := Int" } GT_Contact(in1 := "触摸屏".内室湿度, in2 := 0)
      Coil( "中间变量".内室湿度正常标志 )
   END_RUNG
   // the same network as SCL:
   IF NOT "AlwaysTRUE" THEN
       "模拟量转换函数"(模拟量输入最小值 := 5530,
                 模拟量输入最大值 := 27648,
                 模拟量输入值 := "内室湿度",
                 物理量最小值 := 0.0,
                 物理量最大值 := 1000.0,
                 物理量校准值 := "触摸屏".内室湿度偏差校准,
                 物理量输出值 => "触摸屏".内室湿度);
   END_IF;
   IF "FirstScan" THEN "触摸屏".内室湿度 := 600; END_IF;
   IF "触摸屏".内室湿度 >= 1000 THEN "触摸屏".内室湿度 := 1000; END_IF;
   "中间变量".内室湿度正常标志 := "触摸屏".内室湿度 > 0;
END_REGION

REGION Network 7: 前部温度
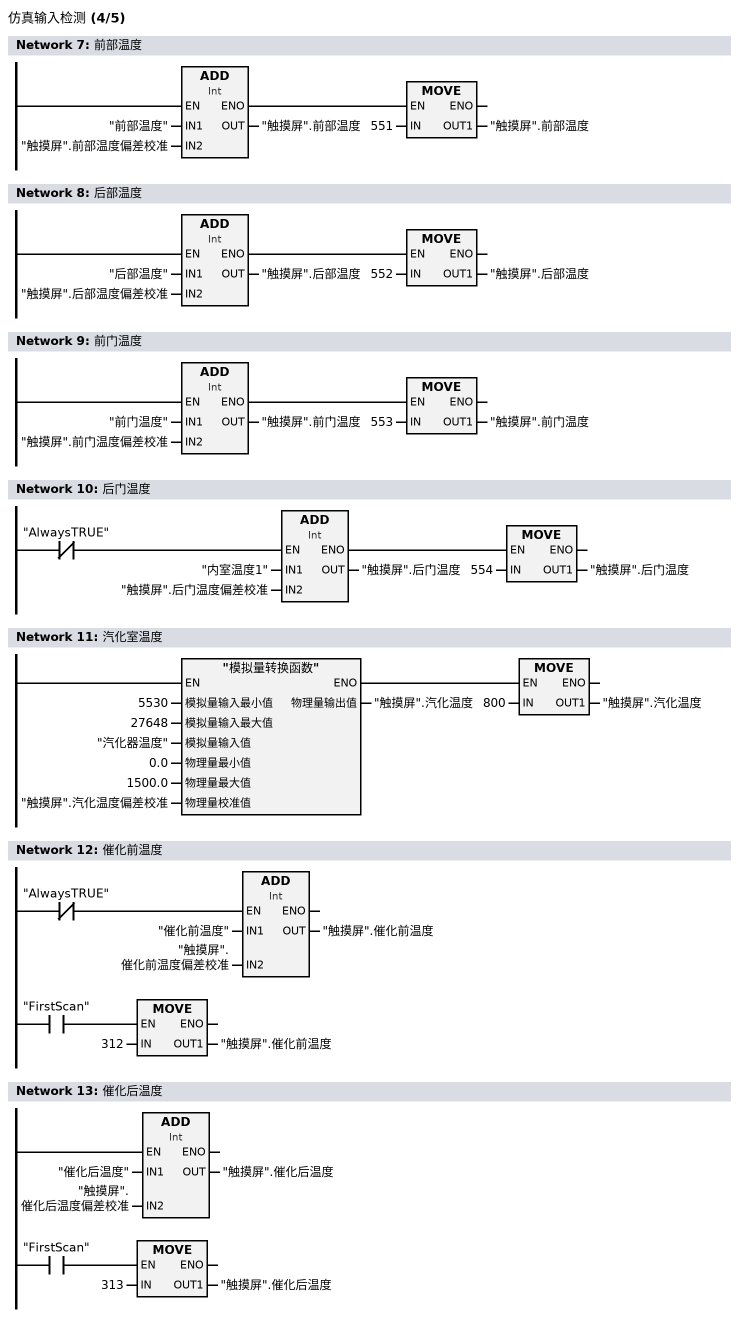
   RUNG wire#powerrail
      { S7_Templates := "SrcType := Int" } Add(in1 := "前部温度", in2 := "触摸屏".前部温度偏差校准, out => "触摸屏".前部温度)
      Move(in := 551, out1 => "触摸屏".前部温度)
   END_RUNG
   // the same network as SCL:
   "触摸屏".前部温度 := "前部温度" + "触摸屏".前部温度偏差校准;
   "触摸屏".前部温度 := 551;
END_REGION

REGION Network 8: 后部温度
   RUNG wire#powerrail
      { S7_Templates := "SrcType := Int" } Add(in1 := "后部温度", in2 := "触摸屏".后部温度偏差校准, out => "触摸屏".后部温度)
      Move(in := 552, out1 => "触摸屏".后部温度)
   END_RUNG
   // the same network as SCL:
   "触摸屏".后部温度 := "后部温度" + "触摸屏".后部温度偏差校准;
   "触摸屏".后部温度 := 552;
END_REGION

REGION Network 9: 前门温度
   RUNG wire#powerrail
      { S7_Templates := "SrcType := Int" } Add(in1 := "前门温度", in2 := "触摸屏".前门温度偏差校准, out => "触摸屏".前门温度)
      Move(in := 553, out1 => "触摸屏".前门温度)
   END_RUNG
   // the same network as SCL:
   "触摸屏".前门温度 := "前门温度" + "触摸屏".前门温度偏差校准;
   "触摸屏".前门温度 := 553;
END_REGION

REGION Network 10: 后门温度
   RUNG wire#powerrail
      I_Contact( "AlwaysTRUE" )
      { S7_Templates := "SrcType := Int" } Add(in1 := "内室温度1", in2 := "触摸屏".后门温度偏差校准, out => "触摸屏".后门温度)
      Move(in := 554, out1 => "触摸屏".后门温度)
   END_RUNG
   // the same network as SCL:
   IF NOT "AlwaysTRUE" THEN
       "触摸屏".后门温度 := "内室温度1" + "触摸屏".后门温度偏差校准;
       "触摸屏".后门温度 := 554;
   END_IF;
END_REGION

REGION Network 11: 汽化室温度
   RUNG wire#powerrail
      "模拟量转换函数"(模拟量输入最小值 := 5530, 模拟量输入最大值 := 27648, 模拟量输入值 := "汽化器温度", 物理量最小值 := 0.0, 物理量最大值 := 1500.0, 物理量校准值 := "触摸屏".汽化温度偏差校准, 物理量输出值 => "触摸屏".汽化温度)
      Move(in := 800, out1 => "触摸屏".汽化温度)
   END_RUNG
   // the same network as SCL:
   "模拟量转换函数"(模拟量输入最小值 := 5530,
             模拟量输入最大值 := 27648,
             模拟量输入值 := "汽化器温度",
             物理量最小值 := 0.0,
             物理量最大值 := 1500.0,
             物理量校准值 := "触摸屏".汽化温度偏差校准,
             物理量输出值 => "触摸屏".汽化温度,
             ENO => #_w1);
   IF #_w1 THEN "触摸屏".汽化温度 := 800; END_IF;
END_REGION

REGION Network 12: 催化前温度
   RUNG wire#powerrail
      I_Contact( "AlwaysTRUE" )
      { S7_Templates := "SrcType := Int" } Add(in1 := "催化前温度", in2 := "触摸屏".催化前温度偏差校准, out => "触摸屏".催化前温度)
   END_RUNG
   RUNG wire#powerrail
      Contact( "FirstScan" )
      Move(in := 312, out1 => "触摸屏".催化前温度)
   END_RUNG
   // the same network as SCL:
   IF NOT "AlwaysTRUE" THEN "触摸屏".催化前温度 := "催化前温度" + "触摸屏".催化前温度偏差校准; END_IF;
   IF "FirstScan" THEN "触摸屏".催化前温度 := 312; END_IF;
END_REGION

REGION Network 13: 催化后温度
   RUNG wire#powerrail
      { S7_Templates := "SrcType := Int" } Add(in1 := "催化后温度", in2 := "触摸屏".催化后温度偏差校准, out => "触摸屏".催化后温度)
   END_RUNG
   RUNG wire#powerrail
      Contact( "FirstScan" )
      Move(in := 313, out1 => "触摸屏".催化后温度)
   END_RUNG
   // the same network as SCL:
   "触摸屏".催化后温度 := "催化后温度" + "触摸屏".催化后温度偏差校准;
   IF "FirstScan" THEN "触摸屏".催化后温度 := 313; END_IF;
END_REGION

REGION Network 14: 每秒更新数据
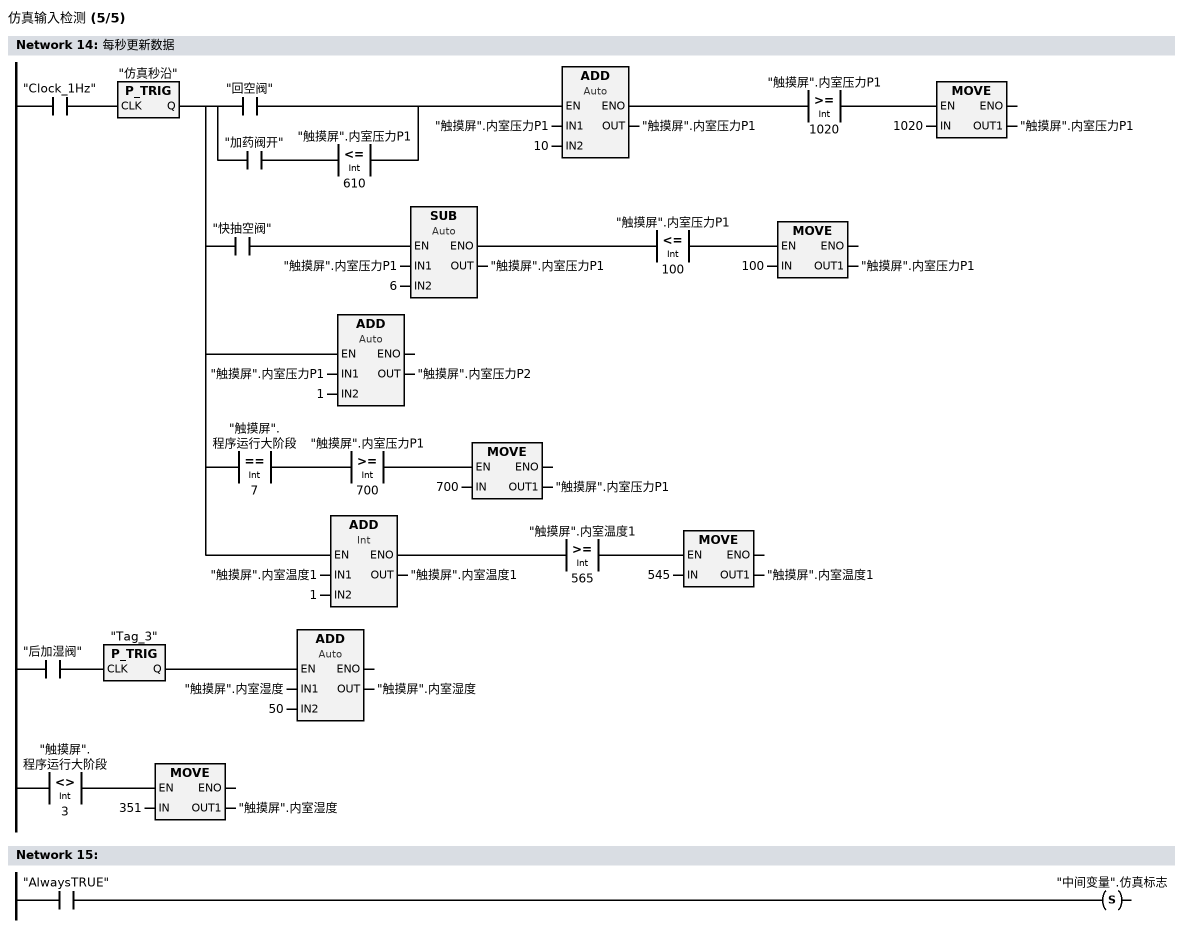
   RUNG wire#powerrail
      Contact( "Clock_1Hz" )
      P_Trig( "仿真秒沿" )
      wire#w1
      Contact( "回空阀" )
      wire#w2
      Add(in1 := "触摸屏".内室压力P1, in2 := 10, out => "触摸屏".内室压力P1)
      { S7_Templates := "SrcType := Int" } GE_Contact(in1 := "触摸屏".内室压力P1, in2 := 1020)
      Move(in := 1020, out1 => "触摸屏".内室压力P1)
   END_RUNG
   RUNG wire#w1
      Contact( "加药阀开" )
      { S7_Templates := "SrcType := Int" } LE_Contact(in1 := "触摸屏".内室压力P1, in2 := 610)
   END_RUNG wire#w2
   RUNG wire#w1
      Contact( "快抽空阀" )
      Sub(in1 := "触摸屏".内室压力P1, in2 := 6, out => "触摸屏".内室压力P1)
      { S7_Templates := "SrcType := Int" } LE_Contact(in1 := "触摸屏".内室压力P1, in2 := 100)
      Move(in := 100, out1 => "触摸屏".内室压力P1)
   END_RUNG
   RUNG wire#w1
      Add(in1 := "触摸屏".内室压力P1, in2 := 1, out => "触摸屏".内室压力P2)
   END_RUNG
   RUNG wire#w1
      { S7_Templates := "SrcType := Int" } EQ_Contact(in1 := "触摸屏".程序运行大阶段, in2 := 7)
      { S7_Templates := "SrcType := Int" } GE_Contact(in1 := "触摸屏".内室压力P1, in2 := 700)
      Move(in := 700, out1 => "触摸屏".内室压力P1)
   END_RUNG
   RUNG wire#w1
      { S7_Templates := "SrcType := Int" } Add(in1 := "触摸屏".内室温度1, in2 := 1, out => "触摸屏".内室温度1)
      { S7_Templates := "SrcType := Int" } GE_Contact(in1 := "触摸屏".内室温度1, in2 := 565)
      Move(in := 545, out1 => "触摸屏".内室温度1)
   END_RUNG
   RUNG wire#powerrail
      Contact( "后加湿阀" )
      P_Trig( "Tag_3" )
      Add(in1 := "触摸屏".内室湿度, in2 := 50, out => "触摸屏".内室湿度)
   END_RUNG
   RUNG wire#powerrail
      { S7_Templates := "SrcType := Int" } NE_Contact(in1 := "触摸屏".程序运行大阶段, in2 := 3)
      Move(in := 351, out1 => "触摸屏".内室湿度)
   END_RUNG
   // the same network as SCL:
   #_w1 := "Clock_1Hz" AND NOT "仿真秒沿";   // rising edge
   "仿真秒沿" := "Clock_1Hz";
   #_w2 := #_w1 AND ("回空阀" OR ("加药阀开" AND ("触摸屏".内室压力P1 <= 610)));
   IF #_w2 THEN "触摸屏".内室压力P1 := "触摸屏".内室压力P1 + 10; END_IF;
   IF #_w2 AND ("触摸屏".内室压力P1 >= 1020) THEN "触摸屏".内室压力P1 := 1020; END_IF;
   #_w3 := #_w1 AND "快抽空阀";
   IF #_w3 THEN "触摸屏".内室压力P1 := "触摸屏".内室压力P1 - 6; END_IF;
   IF #_w3 AND ("触摸屏".内室压力P1 <= 100) THEN "触摸屏".内室压力P1 := 100; END_IF;
   IF #_w1 THEN "触摸屏".内室压力P2 := "触摸屏".内室压力P1 + 1; END_IF;
   IF #_w1 AND ("触摸屏".程序运行大阶段 = 7) AND ("触摸屏".内室压力P1 >= 700) THEN "触摸屏".内室压力P1 := 700; END_IF;
   IF #_w1 THEN "触摸屏".内室温度1 := "触摸屏".内室温度1 + 1; END_IF;
   IF #_w1 AND ("触摸屏".内室温度1 >= 565) THEN "触摸屏".内室温度1 := 545; END_IF;
   #_w4 := "后加湿阀" AND NOT "Tag_3";   // rising edge
   "Tag_3" := "后加湿阀";
   IF #_w4 THEN "触摸屏".内室湿度 := "触摸屏".内室湿度 + 50; END_IF;
   IF "触摸屏".程序运行大阶段 <> 3 THEN "触摸屏".内室湿度 := 351; END_IF;
END_REGION

REGION Network 15
   RUNG wire#powerrail
      Contact( "AlwaysTRUE" )
      S_Coil( "中间变量".仿真标志 )
   END_RUNG
   // the same network as SCL:
   IF "AlwaysTRUE" THEN "中间变量".仿真标志 := TRUE; END_IF;
END_REGION
END_FUNCTION

// folder: 9程序运行控制流程

FUNCTION_BLOCK "8结束"   // FB12, LAD
{ S7_Optimized_Access := 'TRUE' }
VERSION : 0.1
   VAR_INPUT
      启动 : Bool;
      本地大气压 : Int;
      程序暂停位 : Bool;
      内室压力 : Int;
      紧急通风完成标志 : Bool;
   END_VAR
   VAR_OUTPUT
      大阶段运行时间分钟 : Int;
      大阶段运行时间秒 : Int;
      小阶段名称 : Int;
      小阶段运行时间分钟 : Int;
      小阶段运行时间秒 : Int;
      结束阶段完成 : Bool;
      回空阀 : Bool;
      紧急情况阶段完成标志 : Bool;
   END_VAR
   VAR
      统计沿1 : Bool;
      统计沿2 : Bool;
      统计沿3 : Bool;
   END_VAR
   VAR RETAIN
      大阶段时间统计沿 : Bool;
      小阶段时间统计沿 : Bool;
      结束满足压力 : Int;
   END_VAR
   VAR_TEMP
      "中间计算-总秒数" : DInt;
   END_VAR
   VAR_TEMP   // added for the SCL form of the ladder/FBD networks
      _w1 : Bool;
   END_VAR
BEGIN

REGION Network 1: 不启动时将变量清零
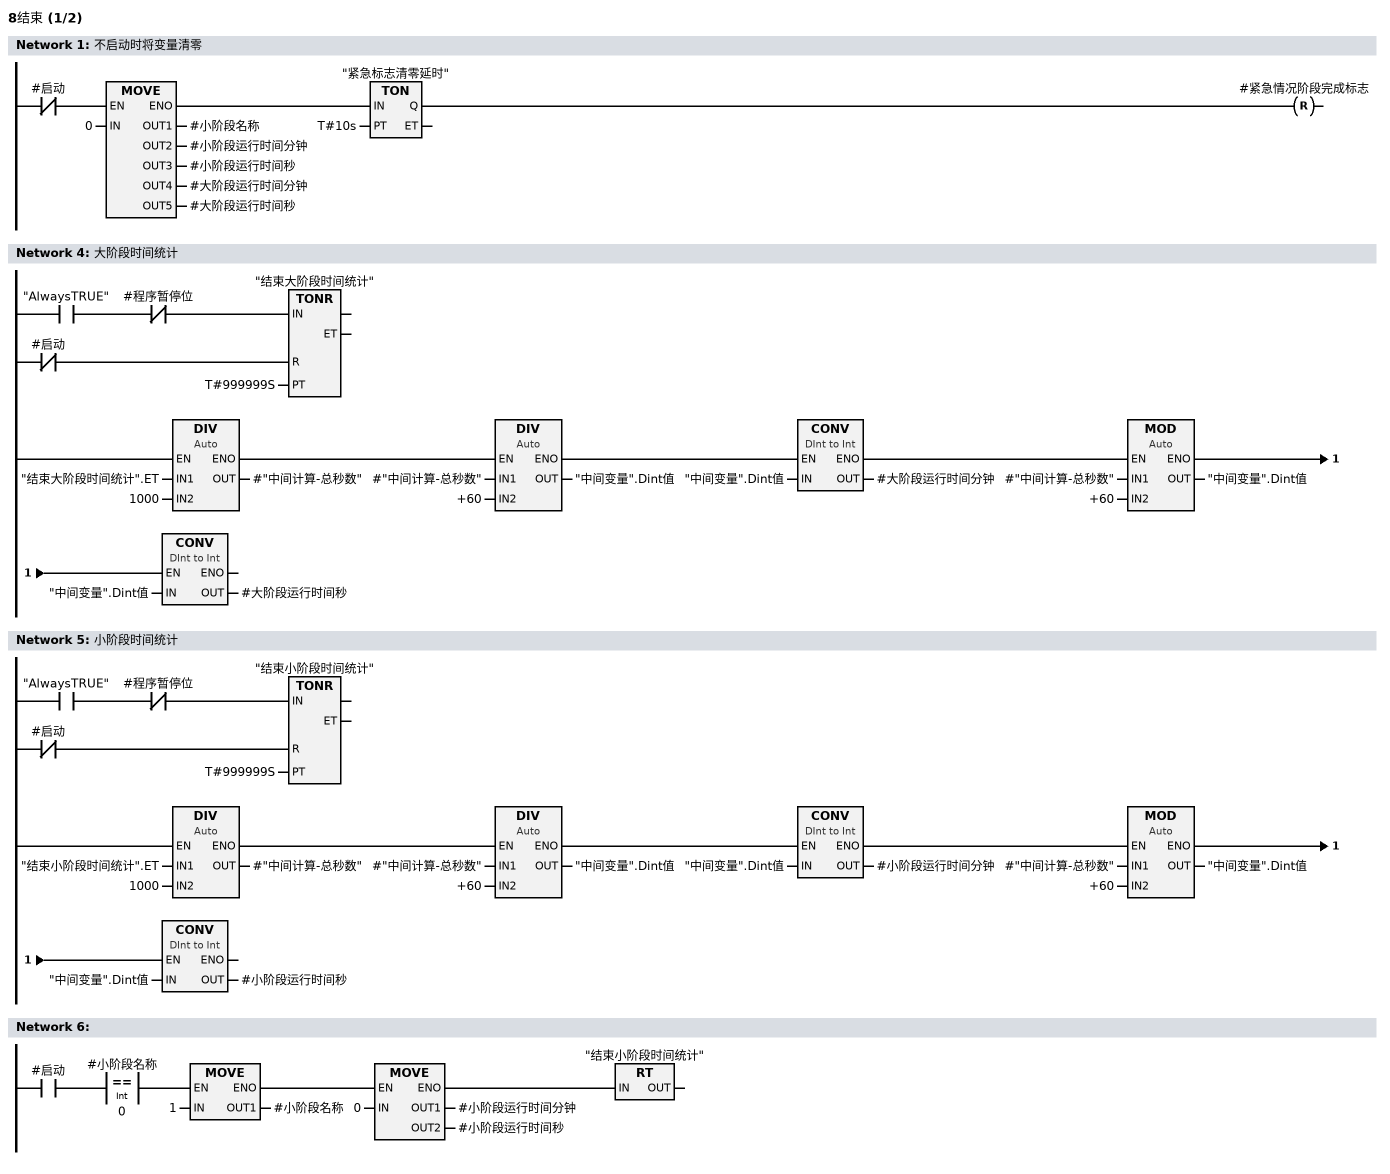
   IF NOT #启动 THEN
       #小阶段名称 := 0;
       #小阶段运行时间分钟 := 0;
       #小阶段运行时间秒 := 0;
       #大阶段运行时间分钟 := 0;
       #大阶段运行时间秒 := 0;
   END_IF;
   "紧急标志清零延时".TON(IN := NOT #启动, PT := T#10s);
   IF "紧急标志清零延时".Q THEN #紧急情况阶段完成标志 := FALSE; END_IF;
END_REGION

REGION Network 4: 大阶段时间统计
   "结束大阶段时间统计".TONR(IN := "AlwaysTRUE" AND NOT #程序暂停位, R := NOT #启动, PT := T#999999S);
   #"中间计算-总秒数" := "结束大阶段时间统计".ET / 1000;
   "中间变量".Dint值 := #"中间计算-总秒数" / +60;
   #大阶段运行时间分钟 := DINT_TO_INT("中间变量".Dint值);
   "中间变量".Dint值 := #"中间计算-总秒数" MOD +60;
   #大阶段运行时间秒 := DINT_TO_INT("中间变量".Dint值);
END_REGION

REGION Network 5: 小阶段时间统计
   "结束小阶段时间统计".TONR(IN := "AlwaysTRUE" AND NOT #程序暂停位, R := NOT #启动, PT := T#999999S);
   #"中间计算-总秒数" := "结束小阶段时间统计".ET / 1000;
   "中间变量".Dint值 := #"中间计算-总秒数" / +60;
   #小阶段运行时间分钟 := DINT_TO_INT("中间变量".Dint值);
   "中间变量".Dint值 := #"中间计算-总秒数" MOD +60;
   #小阶段运行时间秒 := DINT_TO_INT("中间变量".Dint值);
END_REGION

REGION Network 6
   RUNG wire#powerrail
      Contact( #启动 )
      { S7_Templates := "SrcType := Int" } EQ_Contact(in1 := #小阶段名称, in2 := 0)
      Move(in := 1, out1 => #小阶段名称)
      Move(in := 0, out1 => #小阶段运行时间分钟, out2 => #小阶段运行时间秒)
      RT_Coil( "结束小阶段时间统计" )
   END_RUNG
   // the same network as SCL:
   #_w1 := #启动 AND (#小阶段名称 = 0);
   IF #_w1 THEN
       #小阶段名称 := 1;
       #小阶段运行时间分钟 := 0;
       #小阶段运行时间秒 := 0;
       RESET_TIMER("结束小阶段时间统计");
   END_IF;
END_REGION

REGION Network 7: 结束控制流程
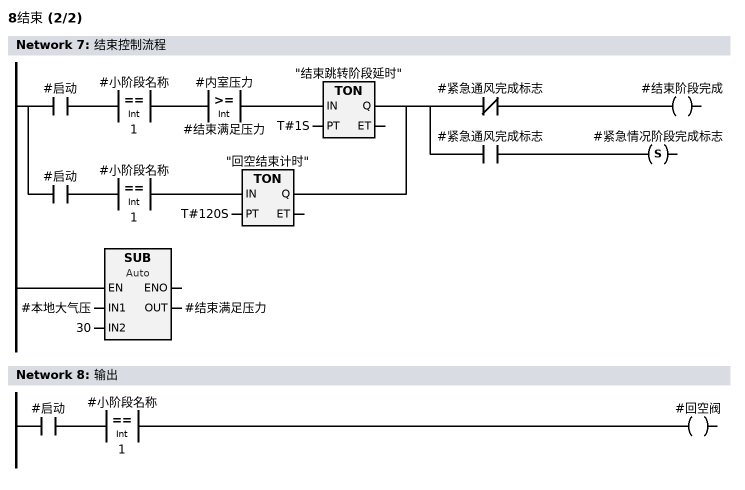
   "结束跳转阶段延时".TON(IN := #启动 AND (#小阶段名称 = 1) AND (#内室压力 >= #结束满足压力), PT := T#1S);
   "回空结束计时".TON(IN := #启动 AND (#小阶段名称 = 1), PT := T#120S);
   #_w1 := "结束跳转阶段延时".Q OR "回空结束计时".Q;
   #结束阶段完成 := #_w1 AND NOT #紧急通风完成标志;
   IF #_w1 AND #紧急通风完成标志 THEN #紧急情况阶段完成标志 := TRUE; END_IF;
   #结束满足压力 := #本地大气压 - 30;
END_REGION

REGION Network 8: 输出
   RUNG wire#powerrail
      Contact( #启动 )
      { S7_Templates := "SrcType := Int" } EQ_Contact(in1 := #小阶段名称, in2 := 1)
      Coil( #回空阀 )
   END_RUNG
   // the same network as SCL:
   #回空阀 := #启动 AND (#小阶段名称 = 1);
END_REGION
END_FUNCTION_BLOCK

FUNCTION_BLOCK "程序倒计时"   // FB13, LAD
{ S7_Optimized_Access := 'TRUE' }
VERSION : 0.1
   VAR
      沿1 : Bool;
      沿2 : Bool;
   END_VAR
   VAR RETAIN
      "预处理时间(秒)" : UInt;
      "预处理时间(分)" : UInt;
      "保压时间(秒)" : UInt;
      "保压时间(分)" : UInt;
      "加湿时间(秒)" : UInt;
      "加湿时间(分)" : UInt;
      "加药时间(秒)" : UInt;
      "加药时间(分)" : UInt;
      "灭菌时间(秒)" : UInt;
      "灭菌时间(分)" : UInt;
      "通风时间(秒)" : UInt;
      "通风时间(分)" : UInt;
      "结束时间(秒)" : UInt;
      "结束时间(分)" : UInt;
      "脉动时间(秒)" : UInt;
      "脉动时间(分)" : UInt;
      总计时间秒 : UInt;
      中间值 : UInt;
   END_VAR
   VAR_TEMP   // added for the SCL form of the ladder/FBD networks
      _w1 : Bool;
      _w2 : Bool;
      _w3 : Bool;
      _w4 : Bool;
      _w5 : Bool;
      _w6 : Bool;
      _w7 : Bool;
      _w8 : Bool;
      _w9 : Bool;
      _w10 : Bool;
      _w11 : Bool;
      _w12 : Bool;
      _w13 : Bool;
      _w14 : Bool;
      _w15 : Bool;
   END_VAR
BEGIN

REGION Network 1: 不运行时间处理
